(* IEC 61131-3 sources: 2026_Projet_YGO_ExcavatriceDragage/TOOLS/TEST_AUTO_CI/RESULTS/L_SIMULATION/reports, 11 files *)

(* ---- FB_Sim_Encoder_test.st ---- *)
(* =======================================================================
   Automated Unit Test - FB_Sim_Encoder
   ======================================================================= *)
TEST 'TC-P13-ENC-001 Enable FALSE conserve la valeur passee par VAR_IN_OUT'
VAR
    fb     : FB_Sim_Encoder;
    rawPos : UDINT := 1000;
END_VAR
    fb.Enable := FALSE;
    fb.StepNumber := 3;
    fb(RawPos := rawPos);
    ASSERT_EQ(fb.RawPosOut, 1000, 'Enable FALSE -> RawPosOut conserve la valeur persistee');
END_TEST

TEST 'TC-P13-ENC-002 Simulation incrementation comptage en montee'
VAR
    fb     : FB_Sim_Encoder;
    rawPos : UDINT := 1000;
    i      : INT;
END_VAR
    fb.Enable := TRUE;
    fb.RelayFwd := TRUE; (* Sens montee *)
    fb.RelayRev := FALSE;
    fb.StepNumber := 3;

    FOR i := 1 TO 10 DO
        fb(RawPos := rawPos);
    END_FOR;

    ASSERT_TRUE(fb.RawPosOut > 1000, 'RelayFwd TRUE -> RawPosOut augmente');
END_TEST

TEST 'TC-P13-034 SpeedReportTauS=0.0 conserve le saut instantane historique (non-regression)'
VAR
    fb     : FB_Sim_Encoder;
    rawPos : UDINT := 1000;
    i      : INT;
END_VAR
    fb.Enable := TRUE;
    fb.RelayFwd := TRUE;
    fb.StepNumber := 5;
    fb.SpeedReportTauS := 0.0;
    FOR i := 1 TO 5 DO
        fb(RawPos := rawPos);
    END_FOR;
    fb.RelayFwd := FALSE;
    fb.CoastDistanceM := 0.0;
    fb(RawPos := rawPos);
    ASSERT_EQ(fb.RawSpdOut, 0, 'Tau=0.0, coupure sans roulis -> vitesse rapportee tombe a 0 des le meme scan');
END_TEST

TEST 'TC-P13-035 SpeedReportTauS>0 fait decroitre RawSpdOut sur plusieurs scans (fidelite AX10, T316)'
VAR
    fb        : FB_Sim_Encoder;
    rawPos    : UDINT := 1000;
    i         : INT;
    spdAtCut  : DINT;
    spdNext   : DINT;
END_VAR
    fb.Enable := TRUE;
    fb.RelayFwd := TRUE;
    fb.StepNumber := 5;
    fb.SpeedReportTauS := 0.15; (* mirror tau M3 identifie sur trace, SYNTHETIQUE treuil *)
    fb.CoastDistanceM := 0.0;
    FOR i := 1 TO 20 DO
        fb(RawPos := rawPos); (* stabilise ReportedSpeedMps a la vitesse palier 5 *)
    END_FOR;
    fb.RelayFwd := FALSE;
    fb(RawPos := rawPos);
    spdAtCut := fb.RawSpdOut;
    fb(RawPos := rawPos);
    spdNext := fb.RawSpdOut;
    ASSERT_TRUE(spdAtCut > 0, 'Coupure relais : vitesse rapportee encore non nulle au 1er scan (pas de saut instantane)');
    ASSERT_TRUE(spdNext < spdAtCut, 'Vitesse rapportee decroit scan apres scan (rampe continue, pas un escalier)');
    ASSERT_TRUE(spdNext > 0, 'Decroissance progressive : pas encore a zero au 2e scan');
END_TEST

TEST 'TC-P13-031 PresetCmd applique PresetValue apres PresetLatencyCycles, mouvement gele pendant la latence'
VAR
    fb     : FB_Sim_Encoder;
    rawPos : UDINT := 1000;
END_VAR
    fb.Enable := TRUE;
    fb.RelayFwd := TRUE; (* commande de mouvement maintenue pendant le preset *)
    fb.StepNumber := 3;
    fb.PresetLatencyCycles := 2;
    fb.PresetValue := 500000;
    fb.PresetCmd := TRUE;
    fb(RawPos := rawPos);
    ASSERT_EQ(fb.RawPosOut, 1000, 'Pendant la latence : position brute conservee, mouvement gele');
    fb(RawPos := rawPos);
    ASSERT_EQ(fb.RawPosOut, 1000, 'Latence non ecoulee : position encore conservee');
    fb(RawPos := rawPos);
    ASSERT_EQ(fb.RawPosOut, 500000, 'Latence ecoulee : PresetValue charge (priorite sur Fwd/Rev)');
END_TEST

TEST 'TC-P13-032 Le comptage descend de facon continue et franchit 0 sans se figer (butee silencieuse supprimee)'
VAR
    fb        : FB_Sim_Encoder;
    rawPos    : UDINT := 41; (* 41 pts : exactement un pas de descente au palier 1 -> atteint 0 au 1er scan *)
    wrapAt41  : UDINT := 4294967255; (* 2^32 - 41 : -41 pts en representation signee 32 bits *)
    wrapAt82  : UDINT := 4294967214; (* 2^32 - 82 : -82 pts *)
END_VAR
    fb.Enable := TRUE;
    fb.RelayRev := TRUE;
    fb.StepNumber := 1; (* 1,0 m/s -> 1,0 x 4096 x 0,010 = 40,96 pts/scan, arrondi a 41 *)
    fb(RawPos := rawPos);
    rawPos := fb.RawPosOut; (* le caller conserve la memoire persistante du codeur *)
    ASSERT_EQ(fb.RawPosOut, 0, 'Un pas de descente amene le comptage exactement a 0 (point de passage)');
    fb(RawPos := rawPos);
    rawPos := fb.RawPosOut;
    ASSERT_TRUE(fb.RawPosOut <> 0, 'Scan suivant : le comptage franchit 0 au lieu de s y figer');
    ASSERT_EQ(fb.RawPosOut, wrapAt41, 'Comptage = -41 pts (aucune borne a 0)');
    fb(RawPos := rawPos);
    ASSERT_EQ(fb.RawPosOut, wrapAt82, 'Le comptage continue de decroitre : -82 pts');
END_TEST

TEST 'TC-P13-036 Comptage a 0 sous commande de descente : le scan suivant ne maintient pas 0'
VAR
    fb       : FB_Sim_Encoder;
    rawPos   : UDINT := 0; (* etat exact du blocage M2 du 2026-09-20 *)
    wrapAt41 : UDINT := 4294967255; (* 2^32 - 41 : -41 pts *)
END_VAR
    fb.Enable := TRUE;
    fb.RelayRev := TRUE;
    fb.StepNumber := 1;
    fb(RawPos := rawPos);
    rawPos := fb.RawPosOut;
    ASSERT_EQ(fb.RawPosOut, wrapAt41, 'Comptage a 0 + descente : passe a -41 pts, ne reste pas bloque a 0');
    fb(RawPos := rawPos);
    ASSERT_EQ(fb.RawPosOut, 4294967214, 'Le comptage poursuit sa descente au scan suivant (-82 pts)');
END_TEST

TEST 'TC-P13-037 Garde de plage : saturation signalee, comptage borne, aucune vitesse publiee'
VAR
    fb         : FB_Sim_Encoder;
    posLimit   : UDINT := 1073741824; (* +2^30 pts : limite de plage du modele *)
    negLimit   : UDINT := 3221225472; (* 2^32 - 2^30 : -2^30 pts en signe *)
END_VAR
    fb.Enable := TRUE;
    fb.RelayFwd := TRUE;
    fb.StepNumber := 5; (* palier 5 : 82 pts/scan *)
    fb(RawPos := posLimit);
    ASSERT_TRUE(fb.CountSaturated, 'Comptage hors plage haute : CountSaturated TRUE (saturation signalee)');
    ASSERT_EQ(fb.RawPosOut, posLimit, 'Comptage borne a la limite de plage (aucun rebouclage UDINT)');
    ASSERT_EQ(fb.RawSpdOut, 0, 'Position bornee : aucune vitesse de mouvement publiee (coherence)');
    fb.RelayFwd := FALSE;
    fb.RelayRev := TRUE;
    fb(RawPos := negLimit);
    ASSERT_TRUE(fb.CountSaturated, 'Comptage hors plage basse : CountSaturated TRUE');
    ASSERT_EQ(fb.RawPosOut, negLimit, 'Comptage borne a la limite basse (aucun rebouclage UDINT)');
    ASSERT_EQ(fb.RawSpdOut, 0, 'Saturation basse : vitesse de mouvement purge');
END_TEST

TEST 'TC-P13-038 Comptage negatif : la montee ramene vers 0 puis au-dela (continuite bidirectionnelle)'
VAR
    fb      : FB_Sim_Encoder;
    rawPos  : UDINT := 4294967255; (* 2^32 - 41 : -41 pts *)
END_VAR
    fb.Enable := TRUE;
    fb.RelayFwd := TRUE;
    fb.RelayRev := FALSE;
    fb.StepNumber := 1;
    fb(RawPos := rawPos);
    rawPos := fb.RawPosOut;
    ASSERT_EQ(fb.RawPosOut, 0, 'Depuis -41 pts : un pas de montee ramene exactement a 0');
    fb(RawPos := rawPos);
    ASSERT_EQ(fb.RawPosOut, 41, 'Le scan suivant poursuit au-dela de 0 (aucune butee dans les deux sens)');
END_TEST

(* ---- FB_Sim_Joystick_test.st ---- *)
(* =======================================================================
   Automated Unit Test - FB_Sim_Joystick
   ======================================================================= *)
TEST 'TC-P13-JOY-001 Enable FALSE -> positionne les axes au neutre (5000)'
VAR
    fb : FB_Sim_Joystick;
END_VAR
    fb.Enable := FALSE;
    fb();
    ASSERT_EQ(fb.RawX, 5000, 'Enable FALSE -> RawX au neutre NeutralRaw=5000');
    ASSERT_EQ(fb.RawY, 5000, 'Enable FALSE -> RawY au neutre NeutralRaw=5000');
    ASSERT_FALSE(fb.RawButton, 'Enable FALSE -> RawButton FALSE');
END_TEST

TEST 'TC-T418-001 Appui avant debattement puis relachement armement'
VAR
    fb : FB_Sim_Joystick;
    i  : INT;
END_VAR
    fb.Enable := TRUE;
    fb(); (* Relachement observe avant nouveau geste *)
    fb.BtnFwd_Up_Close := TRUE;
    fb();
    ASSERT_TRUE(fb.RawButton, 'Appui armement en premier');
    ASSERT_EQ(fb.RawY, 5000, 'Manche au neutre pendant appui');
    ADVANCE_TIME(10000000);
        fb();
ADVANCE_TIME(10000000);
        fb();
ADVANCE_TIME(10000000);
        fb();
ADVANCE_TIME(10000000);
        fb();
ADVANCE_TIME(10000000);
        fb();
ADVANCE_TIME(10000000);
        fb();
ADVANCE_TIME(10000000);
        fb();
ADVANCE_TIME(10000000);
        fb();
ADVANCE_TIME(10000000);
        fb();
ADVANCE_TIME(10000000);
        fb();
    ASSERT_TRUE(fb.RawButton, 'Appui tenu 100 ms');
    ASSERT_EQ(fb.RawY, 5000, 'Aucun debattement avant 200 ms');
    ADVANCE_TIME(10000000);
        fb();
ADVANCE_TIME(10000000);
        fb();
ADVANCE_TIME(10000000);
        fb();
ADVANCE_TIME(10000000);
        fb();
ADVANCE_TIME(10000000);
        fb();
ADVANCE_TIME(10000000);
        fb();
ADVANCE_TIME(10000000);
        fb();
ADVANCE_TIME(10000000);
        fb();
ADVANCE_TIME(10000000);
        fb();
ADVANCE_TIME(10000000);
        fb();
ADVANCE_TIME(10000000);
        fb();
ADVANCE_TIME(10000000);
        fb();
ADVANCE_TIME(10000000);
        fb();
ADVANCE_TIME(10000000);
        fb();
ADVANCE_TIME(10000000);
        fb();
ADVANCE_TIME(10000000);
        fb();
ADVANCE_TIME(10000000);
        fb();
ADVANCE_TIME(10000000);
        fb();
ADVANCE_TIME(10000000);
        fb();
ADVANCE_TIME(10000000);
        fb();
ADVANCE_TIME(10000000);
        fb();
ADVANCE_TIME(10000000);
        fb();
ADVANCE_TIME(10000000);
        fb();
ADVANCE_TIME(10000000);
        fb();
ADVANCE_TIME(10000000);
        fb();
    ASSERT_TRUE(fb.RawY > 5000, 'BtnFwd -> RawY monte vers MaxRaw');
    ASSERT_TRUE(fb.RawButton, 'Armement encore tenu au debut debattement');
    ADVANCE_TIME(10000000);
        fb();
        ASSERT_FALSE(fb.RawButton AND 1 > 20, 'Pas de nouvel appui apres relachement');
ADVANCE_TIME(10000000);
        fb();
        ASSERT_FALSE(fb.RawButton AND 2 > 20, 'Pas de nouvel appui apres relachement');
ADVANCE_TIME(10000000);
        fb();
        ASSERT_FALSE(fb.RawButton AND 3 > 20, 'Pas de nouvel appui apres relachement');
ADVANCE_TIME(10000000);
        fb();
        ASSERT_FALSE(fb.RawButton AND 4 > 20, 'Pas de nouvel appui apres relachement');
ADVANCE_TIME(10000000);
        fb();
        ASSERT_FALSE(fb.RawButton AND 5 > 20, 'Pas de nouvel appui apres relachement');
ADVANCE_TIME(10000000);
        fb();
        ASSERT_FALSE(fb.RawButton AND 6 > 20, 'Pas de nouvel appui apres relachement');
ADVANCE_TIME(10000000);
        fb();
        ASSERT_FALSE(fb.RawButton AND 7 > 20, 'Pas de nouvel appui apres relachement');
ADVANCE_TIME(10000000);
        fb();
        ASSERT_FALSE(fb.RawButton AND 8 > 20, 'Pas de nouvel appui apres relachement');
ADVANCE_TIME(10000000);
        fb();
        ASSERT_FALSE(fb.RawButton AND 9 > 20, 'Pas de nouvel appui apres relachement');
ADVANCE_TIME(10000000);
        fb();
        ASSERT_FALSE(fb.RawButton AND 10 > 20, 'Pas de nouvel appui apres relachement');
ADVANCE_TIME(10000000);
        fb();
        ASSERT_FALSE(fb.RawButton AND 11 > 20, 'Pas de nouvel appui apres relachement');
ADVANCE_TIME(10000000);
        fb();
        ASSERT_FALSE(fb.RawButton AND 12 > 20, 'Pas de nouvel appui apres relachement');
ADVANCE_TIME(10000000);
        fb();
        ASSERT_FALSE(fb.RawButton AND 13 > 20, 'Pas de nouvel appui apres relachement');
ADVANCE_TIME(10000000);
        fb();
        ASSERT_FALSE(fb.RawButton AND 14 > 20, 'Pas de nouvel appui apres relachement');
ADVANCE_TIME(10000000);
        fb();
        ASSERT_FALSE(fb.RawButton AND 15 > 20, 'Pas de nouvel appui apres relachement');
ADVANCE_TIME(10000000);
        fb();
        ASSERT_FALSE(fb.RawButton AND 16 > 20, 'Pas de nouvel appui apres relachement');
ADVANCE_TIME(10000000);
        fb();
        ASSERT_FALSE(fb.RawButton AND 17 > 20, 'Pas de nouvel appui apres relachement');
ADVANCE_TIME(10000000);
        fb();
        ASSERT_FALSE(fb.RawButton AND 18 > 20, 'Pas de nouvel appui apres relachement');
ADVANCE_TIME(10000000);
        fb();
        ASSERT_FALSE(fb.RawButton AND 19 > 20, 'Pas de nouvel appui apres relachement');
ADVANCE_TIME(10000000);
        fb();
        ASSERT_FALSE(fb.RawButton AND 20 > 20, 'Pas de nouvel appui apres relachement');
ADVANCE_TIME(10000000);
        fb();
        ASSERT_FALSE(fb.RawButton AND 21 > 20, 'Pas de nouvel appui apres relachement');
ADVANCE_TIME(10000000);
        fb();
        ASSERT_FALSE(fb.RawButton AND 22 > 20, 'Pas de nouvel appui apres relachement');
ADVANCE_TIME(10000000);
        fb();
        ASSERT_FALSE(fb.RawButton AND 23 > 20, 'Pas de nouvel appui apres relachement');
ADVANCE_TIME(10000000);
        fb();
        ASSERT_FALSE(fb.RawButton AND 24 > 20, 'Pas de nouvel appui apres relachement');
ADVANCE_TIME(10000000);
        fb();
        ASSERT_FALSE(fb.RawButton AND 25 > 20, 'Pas de nouvel appui apres relachement');
ADVANCE_TIME(10000000);
        fb();
        ASSERT_FALSE(fb.RawButton AND 26 > 20, 'Pas de nouvel appui apres relachement');
ADVANCE_TIME(10000000);
        fb();
        ASSERT_FALSE(fb.RawButton AND 27 > 20, 'Pas de nouvel appui apres relachement');
ADVANCE_TIME(10000000);
        fb();
        ASSERT_FALSE(fb.RawButton AND 28 > 20, 'Pas de nouvel appui apres relachement');
ADVANCE_TIME(10000000);
        fb();
        ASSERT_FALSE(fb.RawButton AND 29 > 20, 'Pas de nouvel appui apres relachement');
ADVANCE_TIME(10000000);
        fb();
        ASSERT_FALSE(fb.RawButton AND 30 > 20, 'Pas de nouvel appui apres relachement');
ADVANCE_TIME(10000000);
        fb();
        ASSERT_FALSE(fb.RawButton AND 31 > 20, 'Pas de nouvel appui apres relachement');
ADVANCE_TIME(10000000);
        fb();
        ASSERT_FALSE(fb.RawButton AND 32 > 20, 'Pas de nouvel appui apres relachement');
ADVANCE_TIME(10000000);
        fb();
        ASSERT_FALSE(fb.RawButton AND 33 > 20, 'Pas de nouvel appui apres relachement');
ADVANCE_TIME(10000000);
        fb();
        ASSERT_FALSE(fb.RawButton AND 34 > 20, 'Pas de nouvel appui apres relachement');
ADVANCE_TIME(10000000);
        fb();
        ASSERT_FALSE(fb.RawButton AND 35 > 20, 'Pas de nouvel appui apres relachement');
ADVANCE_TIME(10000000);
        fb();
        ASSERT_FALSE(fb.RawButton AND 36 > 20, 'Pas de nouvel appui apres relachement');
ADVANCE_TIME(10000000);
        fb();
        ASSERT_FALSE(fb.RawButton AND 37 > 20, 'Pas de nouvel appui apres relachement');
ADVANCE_TIME(10000000);
        fb();
        ASSERT_FALSE(fb.RawButton AND 38 > 20, 'Pas de nouvel appui apres relachement');
ADVANCE_TIME(10000000);
        fb();
        ASSERT_FALSE(fb.RawButton AND 39 > 20, 'Pas de nouvel appui apres relachement');
ADVANCE_TIME(10000000);
        fb();
        ASSERT_FALSE(fb.RawButton AND 40 > 20, 'Pas de nouvel appui apres relachement');
ADVANCE_TIME(10000000);
        fb();
        ASSERT_FALSE(fb.RawButton AND 41 > 20, 'Pas de nouvel appui apres relachement');
ADVANCE_TIME(10000000);
        fb();
        ASSERT_FALSE(fb.RawButton AND 42 > 20, 'Pas de nouvel appui apres relachement');
ADVANCE_TIME(10000000);
        fb();
        ASSERT_FALSE(fb.RawButton AND 43 > 20, 'Pas de nouvel appui apres relachement');
ADVANCE_TIME(10000000);
        fb();
        ASSERT_FALSE(fb.RawButton AND 44 > 20, 'Pas de nouvel appui apres relachement');
ADVANCE_TIME(10000000);
        fb();
        ASSERT_FALSE(fb.RawButton AND 45 > 20, 'Pas de nouvel appui apres relachement');
ADVANCE_TIME(10000000);
        fb();
        ASSERT_FALSE(fb.RawButton AND 46 > 20, 'Pas de nouvel appui apres relachement');
ADVANCE_TIME(10000000);
        fb();
        ASSERT_FALSE(fb.RawButton AND 47 > 20, 'Pas de nouvel appui apres relachement');
ADVANCE_TIME(10000000);
        fb();
        ASSERT_FALSE(fb.RawButton AND 48 > 20, 'Pas de nouvel appui apres relachement');
ADVANCE_TIME(10000000);
        fb();
        ASSERT_FALSE(fb.RawButton AND 49 > 20, 'Pas de nouvel appui apres relachement');
ADVANCE_TIME(10000000);
        fb();
        ASSERT_FALSE(fb.RawButton AND 50 > 20, 'Pas de nouvel appui apres relachement');
ADVANCE_TIME(10000000);
        fb();
        ASSERT_FALSE(fb.RawButton AND 51 > 20, 'Pas de nouvel appui apres relachement');
ADVANCE_TIME(10000000);
        fb();
        ASSERT_FALSE(fb.RawButton AND 52 > 20, 'Pas de nouvel appui apres relachement');
ADVANCE_TIME(10000000);
        fb();
        ASSERT_FALSE(fb.RawButton AND 53 > 20, 'Pas de nouvel appui apres relachement');
ADVANCE_TIME(10000000);
        fb();
        ASSERT_FALSE(fb.RawButton AND 54 > 20, 'Pas de nouvel appui apres relachement');
ADVANCE_TIME(10000000);
        fb();
        ASSERT_FALSE(fb.RawButton AND 55 > 20, 'Pas de nouvel appui apres relachement');
ADVANCE_TIME(10000000);
        fb();
        ASSERT_FALSE(fb.RawButton AND 56 > 20, 'Pas de nouvel appui apres relachement');
ADVANCE_TIME(10000000);
        fb();
        ASSERT_FALSE(fb.RawButton AND 57 > 20, 'Pas de nouvel appui apres relachement');
ADVANCE_TIME(10000000);
        fb();
        ASSERT_FALSE(fb.RawButton AND 58 > 20, 'Pas de nouvel appui apres relachement');
ADVANCE_TIME(10000000);
        fb();
        ASSERT_FALSE(fb.RawButton AND 59 > 20, 'Pas de nouvel appui apres relachement');
ADVANCE_TIME(10000000);
        fb();
        ASSERT_FALSE(fb.RawButton AND 60 > 20, 'Pas de nouvel appui apres relachement');
ADVANCE_TIME(10000000);
        fb();
        ASSERT_FALSE(fb.RawButton AND 61 > 20, 'Pas de nouvel appui apres relachement');
ADVANCE_TIME(10000000);
        fb();
        ASSERT_FALSE(fb.RawButton AND 62 > 20, 'Pas de nouvel appui apres relachement');
ADVANCE_TIME(10000000);
        fb();
        ASSERT_FALSE(fb.RawButton AND 63 > 20, 'Pas de nouvel appui apres relachement');
ADVANCE_TIME(10000000);
        fb();
        ASSERT_FALSE(fb.RawButton AND 64 > 20, 'Pas de nouvel appui apres relachement');
ADVANCE_TIME(10000000);
        fb();
        ASSERT_FALSE(fb.RawButton AND 65 > 20, 'Pas de nouvel appui apres relachement');
ADVANCE_TIME(10000000);
        fb();
        ASSERT_FALSE(fb.RawButton AND 66 > 20, 'Pas de nouvel appui apres relachement');
ADVANCE_TIME(10000000);
        fb();
        ASSERT_FALSE(fb.RawButton AND 67 > 20, 'Pas de nouvel appui apres relachement');
ADVANCE_TIME(10000000);
        fb();
        ASSERT_FALSE(fb.RawButton AND 68 > 20, 'Pas de nouvel appui apres relachement');
ADVANCE_TIME(10000000);
        fb();
        ASSERT_FALSE(fb.RawButton AND 69 > 20, 'Pas de nouvel appui apres relachement');
ADVANCE_TIME(10000000);
        fb();
        ASSERT_FALSE(fb.RawButton AND 70 > 20, 'Pas de nouvel appui apres relachement');
ADVANCE_TIME(10000000);
        fb();
        ASSERT_FALSE(fb.RawButton AND 71 > 20, 'Pas de nouvel appui apres relachement');
ADVANCE_TIME(10000000);
        fb();
        ASSERT_FALSE(fb.RawButton AND 72 > 20, 'Pas de nouvel appui apres relachement');
ADVANCE_TIME(10000000);
        fb();
        ASSERT_FALSE(fb.RawButton AND 73 > 20, 'Pas de nouvel appui apres relachement');
ADVANCE_TIME(10000000);
        fb();
        ASSERT_FALSE(fb.RawButton AND 74 > 20, 'Pas de nouvel appui apres relachement');
ADVANCE_TIME(10000000);
        fb();
        ASSERT_FALSE(fb.RawButton AND 75 > 20, 'Pas de nouvel appui apres relachement');
ADVANCE_TIME(10000000);
        fb();
        ASSERT_FALSE(fb.RawButton AND 76 > 20, 'Pas de nouvel appui apres relachement');
ADVANCE_TIME(10000000);
        fb();
        ASSERT_FALSE(fb.RawButton AND 77 > 20, 'Pas de nouvel appui apres relachement');
ADVANCE_TIME(10000000);
        fb();
        ASSERT_FALSE(fb.RawButton AND 78 > 20, 'Pas de nouvel appui apres relachement');
ADVANCE_TIME(10000000);
        fb();
        ASSERT_FALSE(fb.RawButton AND 79 > 20, 'Pas de nouvel appui apres relachement');
ADVANCE_TIME(10000000);
        fb();
        ASSERT_FALSE(fb.RawButton AND 80 > 20, 'Pas de nouvel appui apres relachement');
ADVANCE_TIME(10000000);
        fb();
        ASSERT_FALSE(fb.RawButton AND 81 > 20, 'Pas de nouvel appui apres relachement');
ADVANCE_TIME(10000000);
        fb();
        ASSERT_FALSE(fb.RawButton AND 82 > 20, 'Pas de nouvel appui apres relachement');
ADVANCE_TIME(10000000);
        fb();
        ASSERT_FALSE(fb.RawButton AND 83 > 20, 'Pas de nouvel appui apres relachement');
ADVANCE_TIME(10000000);
        fb();
        ASSERT_FALSE(fb.RawButton AND 84 > 20, 'Pas de nouvel appui apres relachement');
ADVANCE_TIME(10000000);
        fb();
        ASSERT_FALSE(fb.RawButton AND 85 > 20, 'Pas de nouvel appui apres relachement');
ADVANCE_TIME(10000000);
        fb();
        ASSERT_FALSE(fb.RawButton AND 86 > 20, 'Pas de nouvel appui apres relachement');
ADVANCE_TIME(10000000);
        fb();
        ASSERT_FALSE(fb.RawButton AND 87 > 20, 'Pas de nouvel appui apres relachement');
ADVANCE_TIME(10000000);
        fb();
        ASSERT_FALSE(fb.RawButton AND 88 > 20, 'Pas de nouvel appui apres relachement');
ADVANCE_TIME(10000000);
        fb();
        ASSERT_FALSE(fb.RawButton AND 89 > 20, 'Pas de nouvel appui apres relachement');
ADVANCE_TIME(10000000);
        fb();
        ASSERT_FALSE(fb.RawButton AND 90 > 20, 'Pas de nouvel appui apres relachement');
ADVANCE_TIME(10000000);
        fb();
        ASSERT_FALSE(fb.RawButton AND 91 > 20, 'Pas de nouvel appui apres relachement');
ADVANCE_TIME(10000000);
        fb();
        ASSERT_FALSE(fb.RawButton AND 92 > 20, 'Pas de nouvel appui apres relachement');
ADVANCE_TIME(10000000);
        fb();
        ASSERT_FALSE(fb.RawButton AND 93 > 20, 'Pas de nouvel appui apres relachement');
ADVANCE_TIME(10000000);
        fb();
        ASSERT_FALSE(fb.RawButton AND 94 > 20, 'Pas de nouvel appui apres relachement');
ADVANCE_TIME(10000000);
        fb();
        ASSERT_FALSE(fb.RawButton AND 95 > 20, 'Pas de nouvel appui apres relachement');
ADVANCE_TIME(10000000);
        fb();
        ASSERT_FALSE(fb.RawButton AND 96 > 20, 'Pas de nouvel appui apres relachement');
ADVANCE_TIME(10000000);
        fb();
        ASSERT_FALSE(fb.RawButton AND 97 > 20, 'Pas de nouvel appui apres relachement');
ADVANCE_TIME(10000000);
        fb();
        ASSERT_FALSE(fb.RawButton AND 98 > 20, 'Pas de nouvel appui apres relachement');
ADVANCE_TIME(10000000);
        fb();
        ASSERT_FALSE(fb.RawButton AND 99 > 20, 'Pas de nouvel appui apres relachement');
ADVANCE_TIME(10000000);
        fb();
        ASSERT_FALSE(fb.RawButton AND 100 > 20, 'Pas de nouvel appui apres relachement');
ADVANCE_TIME(10000000);
        fb();
        ASSERT_FALSE(fb.RawButton AND 101 > 20, 'Pas de nouvel appui apres relachement');
ADVANCE_TIME(10000000);
        fb();
        ASSERT_FALSE(fb.RawButton AND 102 > 20, 'Pas de nouvel appui apres relachement');
ADVANCE_TIME(10000000);
        fb();
        ASSERT_FALSE(fb.RawButton AND 103 > 20, 'Pas de nouvel appui apres relachement');
ADVANCE_TIME(10000000);
        fb();
        ASSERT_FALSE(fb.RawButton AND 104 > 20, 'Pas de nouvel appui apres relachement');
ADVANCE_TIME(10000000);
        fb();
        ASSERT_FALSE(fb.RawButton AND 105 > 20, 'Pas de nouvel appui apres relachement');
ADVANCE_TIME(10000000);
        fb();
        ASSERT_FALSE(fb.RawButton AND 106 > 20, 'Pas de nouvel appui apres relachement');
ADVANCE_TIME(10000000);
        fb();
        ASSERT_FALSE(fb.RawButton AND 107 > 20, 'Pas de nouvel appui apres relachement');
ADVANCE_TIME(10000000);
        fb();
        ASSERT_FALSE(fb.RawButton AND 108 > 20, 'Pas de nouvel appui apres relachement');
ADVANCE_TIME(10000000);
        fb();
        ASSERT_FALSE(fb.RawButton AND 109 > 20, 'Pas de nouvel appui apres relachement');
ADVANCE_TIME(10000000);
        fb();
        ASSERT_FALSE(fb.RawButton AND 110 > 20, 'Pas de nouvel appui apres relachement');
ADVANCE_TIME(10000000);
        fb();
        ASSERT_FALSE(fb.RawButton AND 111 > 20, 'Pas de nouvel appui apres relachement');
ADVANCE_TIME(10000000);
        fb();
        ASSERT_FALSE(fb.RawButton AND 112 > 20, 'Pas de nouvel appui apres relachement');
ADVANCE_TIME(10000000);
        fb();
        ASSERT_FALSE(fb.RawButton AND 113 > 20, 'Pas de nouvel appui apres relachement');
ADVANCE_TIME(10000000);
        fb();
        ASSERT_FALSE(fb.RawButton AND 114 > 20, 'Pas de nouvel appui apres relachement');
ADVANCE_TIME(10000000);
        fb();
        ASSERT_FALSE(fb.RawButton AND 115 > 20, 'Pas de nouvel appui apres relachement');
ADVANCE_TIME(10000000);
        fb();
        ASSERT_FALSE(fb.RawButton AND 116 > 20, 'Pas de nouvel appui apres relachement');
ADVANCE_TIME(10000000);
        fb();
        ASSERT_FALSE(fb.RawButton AND 117 > 20, 'Pas de nouvel appui apres relachement');
ADVANCE_TIME(10000000);
        fb();
        ASSERT_FALSE(fb.RawButton AND 118 > 20, 'Pas de nouvel appui apres relachement');
ADVANCE_TIME(10000000);
        fb();
        ASSERT_FALSE(fb.RawButton AND 119 > 20, 'Pas de nouvel appui apres relachement');
ADVANCE_TIME(10000000);
        fb();
        ASSERT_FALSE(fb.RawButton AND 120 > 20, 'Pas de nouvel appui apres relachement');
ADVANCE_TIME(10000000);
        fb();
        ASSERT_FALSE(fb.RawButton AND 121 > 20, 'Pas de nouvel appui apres relachement');
ADVANCE_TIME(10000000);
        fb();
        ASSERT_FALSE(fb.RawButton AND 122 > 20, 'Pas de nouvel appui apres relachement');
ADVANCE_TIME(10000000);
        fb();
        ASSERT_FALSE(fb.RawButton AND 123 > 20, 'Pas de nouvel appui apres relachement');
ADVANCE_TIME(10000000);
        fb();
        ASSERT_FALSE(fb.RawButton AND 124 > 20, 'Pas de nouvel appui apres relachement');
ADVANCE_TIME(10000000);
        fb();
        ASSERT_FALSE(fb.RawButton AND 125 > 20, 'Pas de nouvel appui apres relachement');
ADVANCE_TIME(10000000);
        fb();
        ASSERT_FALSE(fb.RawButton AND 126 > 20, 'Pas de nouvel appui apres relachement');
ADVANCE_TIME(10000000);
        fb();
        ASSERT_FALSE(fb.RawButton AND 127 > 20, 'Pas de nouvel appui apres relachement');
ADVANCE_TIME(10000000);
        fb();
        ASSERT_FALSE(fb.RawButton AND 128 > 20, 'Pas de nouvel appui apres relachement');
ADVANCE_TIME(10000000);
        fb();
        ASSERT_FALSE(fb.RawButton AND 129 > 20, 'Pas de nouvel appui apres relachement');
ADVANCE_TIME(10000000);
        fb();
        ASSERT_FALSE(fb.RawButton AND 130 > 20, 'Pas de nouvel appui apres relachement');
ADVANCE_TIME(10000000);
        fb();
        ASSERT_FALSE(fb.RawButton AND 131 > 20, 'Pas de nouvel appui apres relachement');
ADVANCE_TIME(10000000);
        fb();
        ASSERT_FALSE(fb.RawButton AND 132 > 20, 'Pas de nouvel appui apres relachement');
ADVANCE_TIME(10000000);
        fb();
        ASSERT_FALSE(fb.RawButton AND 133 > 20, 'Pas de nouvel appui apres relachement');
ADVANCE_TIME(10000000);
        fb();
        ASSERT_FALSE(fb.RawButton AND 134 > 20, 'Pas de nouvel appui apres relachement');
ADVANCE_TIME(10000000);
        fb();
        ASSERT_FALSE(fb.RawButton AND 135 > 20, 'Pas de nouvel appui apres relachement');
ADVANCE_TIME(10000000);
        fb();
        ASSERT_FALSE(fb.RawButton AND 136 > 20, 'Pas de nouvel appui apres relachement');
ADVANCE_TIME(10000000);
        fb();
        ASSERT_FALSE(fb.RawButton AND 137 > 20, 'Pas de nouvel appui apres relachement');
ADVANCE_TIME(10000000);
        fb();
        ASSERT_FALSE(fb.RawButton AND 138 > 20, 'Pas de nouvel appui apres relachement');
ADVANCE_TIME(10000000);
        fb();
        ASSERT_FALSE(fb.RawButton AND 139 > 20, 'Pas de nouvel appui apres relachement');
ADVANCE_TIME(10000000);
        fb();
        ASSERT_FALSE(fb.RawButton AND 140 > 20, 'Pas de nouvel appui apres relachement');
ADVANCE_TIME(10000000);
        fb();
        ASSERT_FALSE(fb.RawButton AND 141 > 20, 'Pas de nouvel appui apres relachement');
ADVANCE_TIME(10000000);
        fb();
        ASSERT_FALSE(fb.RawButton AND 142 > 20, 'Pas de nouvel appui apres relachement');
ADVANCE_TIME(10000000);
        fb();
        ASSERT_FALSE(fb.RawButton AND 143 > 20, 'Pas de nouvel appui apres relachement');
ADVANCE_TIME(10000000);
        fb();
        ASSERT_FALSE(fb.RawButton AND 144 > 20, 'Pas de nouvel appui apres relachement');
ADVANCE_TIME(10000000);
        fb();
        ASSERT_FALSE(fb.RawButton AND 145 > 20, 'Pas de nouvel appui apres relachement');
ADVANCE_TIME(10000000);
        fb();
        ASSERT_FALSE(fb.RawButton AND 146 > 20, 'Pas de nouvel appui apres relachement');
ADVANCE_TIME(10000000);
        fb();
        ASSERT_FALSE(fb.RawButton AND 147 > 20, 'Pas de nouvel appui apres relachement');
ADVANCE_TIME(10000000);
        fb();
        ASSERT_FALSE(fb.RawButton AND 148 > 20, 'Pas de nouvel appui apres relachement');
ADVANCE_TIME(10000000);
        fb();
        ASSERT_FALSE(fb.RawButton AND 149 > 20, 'Pas de nouvel appui apres relachement');
ADVANCE_TIME(10000000);
        fb();
        ASSERT_FALSE(fb.RawButton AND 150 > 20, 'Pas de nouvel appui apres relachement');
ADVANCE_TIME(10000000);
        fb();
        ASSERT_FALSE(fb.RawButton AND 151 > 20, 'Pas de nouvel appui apres relachement');
ADVANCE_TIME(10000000);
        fb();
        ASSERT_FALSE(fb.RawButton AND 152 > 20, 'Pas de nouvel appui apres relachement');
ADVANCE_TIME(10000000);
        fb();
        ASSERT_FALSE(fb.RawButton AND 153 > 20, 'Pas de nouvel appui apres relachement');
ADVANCE_TIME(10000000);
        fb();
        ASSERT_FALSE(fb.RawButton AND 154 > 20, 'Pas de nouvel appui apres relachement');
ADVANCE_TIME(10000000);
        fb();
        ASSERT_FALSE(fb.RawButton AND 155 > 20, 'Pas de nouvel appui apres relachement');
ADVANCE_TIME(10000000);
        fb();
        ASSERT_FALSE(fb.RawButton AND 156 > 20, 'Pas de nouvel appui apres relachement');
ADVANCE_TIME(10000000);
        fb();
        ASSERT_FALSE(fb.RawButton AND 157 > 20, 'Pas de nouvel appui apres relachement');
ADVANCE_TIME(10000000);
        fb();
        ASSERT_FALSE(fb.RawButton AND 158 > 20, 'Pas de nouvel appui apres relachement');
ADVANCE_TIME(10000000);
        fb();
        ASSERT_FALSE(fb.RawButton AND 159 > 20, 'Pas de nouvel appui apres relachement');
ADVANCE_TIME(10000000);
        fb();
        ASSERT_FALSE(fb.RawButton AND 160 > 20, 'Pas de nouvel appui apres relachement');
ADVANCE_TIME(10000000);
        fb();
        ASSERT_FALSE(fb.RawButton AND 161 > 20, 'Pas de nouvel appui apres relachement');
ADVANCE_TIME(10000000);
        fb();
        ASSERT_FALSE(fb.RawButton AND 162 > 20, 'Pas de nouvel appui apres relachement');
ADVANCE_TIME(10000000);
        fb();
        ASSERT_FALSE(fb.RawButton AND 163 > 20, 'Pas de nouvel appui apres relachement');
ADVANCE_TIME(10000000);
        fb();
        ASSERT_FALSE(fb.RawButton AND 164 > 20, 'Pas de nouvel appui apres relachement');
ADVANCE_TIME(10000000);
        fb();
        ASSERT_FALSE(fb.RawButton AND 165 > 20, 'Pas de nouvel appui apres relachement');
ADVANCE_TIME(10000000);
        fb();
        ASSERT_FALSE(fb.RawButton AND 166 > 20, 'Pas de nouvel appui apres relachement');
ADVANCE_TIME(10000000);
        fb();
        ASSERT_FALSE(fb.RawButton AND 167 > 20, 'Pas de nouvel appui apres relachement');
ADVANCE_TIME(10000000);
        fb();
        ASSERT_FALSE(fb.RawButton AND 168 > 20, 'Pas de nouvel appui apres relachement');
ADVANCE_TIME(10000000);
        fb();
        ASSERT_FALSE(fb.RawButton AND 169 > 20, 'Pas de nouvel appui apres relachement');
ADVANCE_TIME(10000000);
        fb();
        ASSERT_FALSE(fb.RawButton AND 170 > 20, 'Pas de nouvel appui apres relachement');
ADVANCE_TIME(10000000);
        fb();
        ASSERT_FALSE(fb.RawButton AND 171 > 20, 'Pas de nouvel appui apres relachement');
ADVANCE_TIME(10000000);
        fb();
        ASSERT_FALSE(fb.RawButton AND 172 > 20, 'Pas de nouvel appui apres relachement');
ADVANCE_TIME(10000000);
        fb();
        ASSERT_FALSE(fb.RawButton AND 173 > 20, 'Pas de nouvel appui apres relachement');
ADVANCE_TIME(10000000);
        fb();
        ASSERT_FALSE(fb.RawButton AND 174 > 20, 'Pas de nouvel appui apres relachement');
ADVANCE_TIME(10000000);
        fb();
        ASSERT_FALSE(fb.RawButton AND 175 > 20, 'Pas de nouvel appui apres relachement');
ADVANCE_TIME(10000000);
        fb();
        ASSERT_FALSE(fb.RawButton AND 176 > 20, 'Pas de nouvel appui apres relachement');
ADVANCE_TIME(10000000);
        fb();
        ASSERT_FALSE(fb.RawButton AND 177 > 20, 'Pas de nouvel appui apres relachement');
ADVANCE_TIME(10000000);
        fb();
        ASSERT_FALSE(fb.RawButton AND 178 > 20, 'Pas de nouvel appui apres relachement');
ADVANCE_TIME(10000000);
        fb();
        ASSERT_FALSE(fb.RawButton AND 179 > 20, 'Pas de nouvel appui apres relachement');
ADVANCE_TIME(10000000);
        fb();
        ASSERT_FALSE(fb.RawButton AND 180 > 20, 'Pas de nouvel appui apres relachement');
ADVANCE_TIME(10000000);
        fb();
        ASSERT_FALSE(fb.RawButton AND 181 > 20, 'Pas de nouvel appui apres relachement');
ADVANCE_TIME(10000000);
        fb();
        ASSERT_FALSE(fb.RawButton AND 182 > 20, 'Pas de nouvel appui apres relachement');
ADVANCE_TIME(10000000);
        fb();
        ASSERT_FALSE(fb.RawButton AND 183 > 20, 'Pas de nouvel appui apres relachement');
ADVANCE_TIME(10000000);
        fb();
        ASSERT_FALSE(fb.RawButton AND 184 > 20, 'Pas de nouvel appui apres relachement');
ADVANCE_TIME(10000000);
        fb();
        ASSERT_FALSE(fb.RawButton AND 185 > 20, 'Pas de nouvel appui apres relachement');
ADVANCE_TIME(10000000);
        fb();
        ASSERT_FALSE(fb.RawButton AND 186 > 20, 'Pas de nouvel appui apres relachement');
ADVANCE_TIME(10000000);
        fb();
        ASSERT_FALSE(fb.RawButton AND 187 > 20, 'Pas de nouvel appui apres relachement');
ADVANCE_TIME(10000000);
        fb();
        ASSERT_FALSE(fb.RawButton AND 188 > 20, 'Pas de nouvel appui apres relachement');
ADVANCE_TIME(10000000);
        fb();
        ASSERT_FALSE(fb.RawButton AND 189 > 20, 'Pas de nouvel appui apres relachement');
ADVANCE_TIME(10000000);
        fb();
        ASSERT_FALSE(fb.RawButton AND 190 > 20, 'Pas de nouvel appui apres relachement');
ADVANCE_TIME(10000000);
        fb();
        ASSERT_FALSE(fb.RawButton AND 191 > 20, 'Pas de nouvel appui apres relachement');
ADVANCE_TIME(10000000);
        fb();
        ASSERT_FALSE(fb.RawButton AND 192 > 20, 'Pas de nouvel appui apres relachement');
ADVANCE_TIME(10000000);
        fb();
        ASSERT_FALSE(fb.RawButton AND 193 > 20, 'Pas de nouvel appui apres relachement');
ADVANCE_TIME(10000000);
        fb();
        ASSERT_FALSE(fb.RawButton AND 194 > 20, 'Pas de nouvel appui apres relachement');
ADVANCE_TIME(10000000);
        fb();
        ASSERT_FALSE(fb.RawButton AND 195 > 20, 'Pas de nouvel appui apres relachement');
ADVANCE_TIME(10000000);
        fb();
        ASSERT_FALSE(fb.RawButton AND 196 > 20, 'Pas de nouvel appui apres relachement');
ADVANCE_TIME(10000000);
        fb();
        ASSERT_FALSE(fb.RawButton AND 197 > 20, 'Pas de nouvel appui apres relachement');
ADVANCE_TIME(10000000);
        fb();
        ASSERT_FALSE(fb.RawButton AND 198 > 20, 'Pas de nouvel appui apres relachement');
ADVANCE_TIME(10000000);
        fb();
        ASSERT_FALSE(fb.RawButton AND 199 > 20, 'Pas de nouvel appui apres relachement');
ADVANCE_TIME(10000000);
        fb();
        ASSERT_FALSE(fb.RawButton AND 200 > 20, 'Pas de nouvel appui apres relachement');
ADVANCE_TIME(10000000);
        fb();
        ASSERT_FALSE(fb.RawButton AND 201 > 20, 'Pas de nouvel appui apres relachement');
ADVANCE_TIME(10000000);
        fb();
        ASSERT_FALSE(fb.RawButton AND 202 > 20, 'Pas de nouvel appui apres relachement');
ADVANCE_TIME(10000000);
        fb();
        ASSERT_FALSE(fb.RawButton AND 203 > 20, 'Pas de nouvel appui apres relachement');
ADVANCE_TIME(10000000);
        fb();
        ASSERT_FALSE(fb.RawButton AND 204 > 20, 'Pas de nouvel appui apres relachement');
ADVANCE_TIME(10000000);
        fb();
        ASSERT_FALSE(fb.RawButton AND 205 > 20, 'Pas de nouvel appui apres relachement');
ADVANCE_TIME(10000000);
        fb();
        ASSERT_FALSE(fb.RawButton AND 206 > 20, 'Pas de nouvel appui apres relachement');
ADVANCE_TIME(10000000);
        fb();
        ASSERT_FALSE(fb.RawButton AND 207 > 20, 'Pas de nouvel appui apres relachement');
ADVANCE_TIME(10000000);
        fb();
        ASSERT_FALSE(fb.RawButton AND 208 > 20, 'Pas de nouvel appui apres relachement');
ADVANCE_TIME(10000000);
        fb();
        ASSERT_FALSE(fb.RawButton AND 209 > 20, 'Pas de nouvel appui apres relachement');
ADVANCE_TIME(10000000);
        fb();
        ASSERT_FALSE(fb.RawButton AND 210 > 20, 'Pas de nouvel appui apres relachement');
ADVANCE_TIME(10000000);
        fb();
        ASSERT_FALSE(fb.RawButton AND 211 > 20, 'Pas de nouvel appui apres relachement');
ADVANCE_TIME(10000000);
        fb();
        ASSERT_FALSE(fb.RawButton AND 212 > 20, 'Pas de nouvel appui apres relachement');
ADVANCE_TIME(10000000);
        fb();
        ASSERT_FALSE(fb.RawButton AND 213 > 20, 'Pas de nouvel appui apres relachement');
ADVANCE_TIME(10000000);
        fb();
        ASSERT_FALSE(fb.RawButton AND 214 > 20, 'Pas de nouvel appui apres relachement');
ADVANCE_TIME(10000000);
        fb();
        ASSERT_FALSE(fb.RawButton AND 215 > 20, 'Pas de nouvel appui apres relachement');
ADVANCE_TIME(10000000);
        fb();
        ASSERT_FALSE(fb.RawButton AND 216 > 20, 'Pas de nouvel appui apres relachement');
ADVANCE_TIME(10000000);
        fb();
        ASSERT_FALSE(fb.RawButton AND 217 > 20, 'Pas de nouvel appui apres relachement');
ADVANCE_TIME(10000000);
        fb();
        ASSERT_FALSE(fb.RawButton AND 218 > 20, 'Pas de nouvel appui apres relachement');
ADVANCE_TIME(10000000);
        fb();
        ASSERT_FALSE(fb.RawButton AND 219 > 20, 'Pas de nouvel appui apres relachement');
ADVANCE_TIME(10000000);
        fb();
        ASSERT_FALSE(fb.RawButton AND 220 > 20, 'Pas de nouvel appui apres relachement');
    ASSERT_FALSE(fb.RawButton, 'Bouton armement relache malgre maintien IHM');
    ASSERT_TRUE(fb.RawY > 9000, 'Manche reste deplace');
    fb.BtnFwd_Up_Close := FALSE;
    ADVANCE_TIME(10000000);
        fb();
ADVANCE_TIME(10000000);
        fb();
ADVANCE_TIME(10000000);
        fb();
ADVANCE_TIME(10000000);
        fb();
ADVANCE_TIME(10000000);
        fb();
ADVANCE_TIME(10000000);
        fb();
ADVANCE_TIME(10000000);
        fb();
ADVANCE_TIME(10000000);
        fb();
ADVANCE_TIME(10000000);
        fb();
ADVANCE_TIME(10000000);
        fb();
ADVANCE_TIME(10000000);
        fb();
ADVANCE_TIME(10000000);
        fb();
ADVANCE_TIME(10000000);
        fb();
ADVANCE_TIME(10000000);
        fb();
ADVANCE_TIME(10000000);
        fb();
ADVANCE_TIME(10000000);
        fb();
ADVANCE_TIME(10000000);
        fb();
ADVANCE_TIME(10000000);
        fb();
ADVANCE_TIME(10000000);
        fb();
ADVANCE_TIME(10000000);
        fb();
ADVANCE_TIME(10000000);
        fb();
ADVANCE_TIME(10000000);
        fb();
ADVANCE_TIME(10000000);
        fb();
ADVANCE_TIME(10000000);
        fb();
ADVANCE_TIME(10000000);
        fb();
ADVANCE_TIME(10000000);
        fb();
ADVANCE_TIME(10000000);
        fb();
ADVANCE_TIME(10000000);
        fb();
ADVANCE_TIME(10000000);
        fb();
ADVANCE_TIME(10000000);
        fb();
    ASSERT_EQ(fb.RawY, 5000, 'Retour au neutre au relachement IHM');
    ASSERT_FALSE(fb.ModelActive, 'Fin de propriete automatique');
END_TEST

TEST 'TC-T418-002 Bouton deja tenu au demarrage ou reactivation'
VAR
    fb : FB_Sim_Joystick;
    i : INT;
END_VAR
    fb.Enable := TRUE; fb.BtnRight_Fwd_MAINT := TRUE;
    ADVANCE_TIME(10000000); fb();
        ASSERT_FALSE(fb.RawButton, 'Demarrage tenu ne simule aucun appui');
        ASSERT_EQ(fb.RawX, 5000, 'Demarrage tenu neutre');
ADVANCE_TIME(10000000); fb();
        ASSERT_FALSE(fb.RawButton, 'Demarrage tenu ne simule aucun appui');
        ASSERT_EQ(fb.RawX, 5000, 'Demarrage tenu neutre');
ADVANCE_TIME(10000000); fb();
        ASSERT_FALSE(fb.RawButton, 'Demarrage tenu ne simule aucun appui');
        ASSERT_EQ(fb.RawX, 5000, 'Demarrage tenu neutre');
ADVANCE_TIME(10000000); fb();
        ASSERT_FALSE(fb.RawButton, 'Demarrage tenu ne simule aucun appui');
        ASSERT_EQ(fb.RawX, 5000, 'Demarrage tenu neutre');
ADVANCE_TIME(10000000); fb();
        ASSERT_FALSE(fb.RawButton, 'Demarrage tenu ne simule aucun appui');
        ASSERT_EQ(fb.RawX, 5000, 'Demarrage tenu neutre');
ADVANCE_TIME(10000000); fb();
        ASSERT_FALSE(fb.RawButton, 'Demarrage tenu ne simule aucun appui');
        ASSERT_EQ(fb.RawX, 5000, 'Demarrage tenu neutre');
ADVANCE_TIME(10000000); fb();
        ASSERT_FALSE(fb.RawButton, 'Demarrage tenu ne simule aucun appui');
        ASSERT_EQ(fb.RawX, 5000, 'Demarrage tenu neutre');
ADVANCE_TIME(10000000); fb();
        ASSERT_FALSE(fb.RawButton, 'Demarrage tenu ne simule aucun appui');
        ASSERT_EQ(fb.RawX, 5000, 'Demarrage tenu neutre');
ADVANCE_TIME(10000000); fb();
        ASSERT_FALSE(fb.RawButton, 'Demarrage tenu ne simule aucun appui');
        ASSERT_EQ(fb.RawX, 5000, 'Demarrage tenu neutre');
ADVANCE_TIME(10000000); fb();
        ASSERT_FALSE(fb.RawButton, 'Demarrage tenu ne simule aucun appui');
        ASSERT_EQ(fb.RawX, 5000, 'Demarrage tenu neutre');
ADVANCE_TIME(10000000); fb();
        ASSERT_FALSE(fb.RawButton, 'Demarrage tenu ne simule aucun appui');
        ASSERT_EQ(fb.RawX, 5000, 'Demarrage tenu neutre');
ADVANCE_TIME(10000000); fb();
        ASSERT_FALSE(fb.RawButton, 'Demarrage tenu ne simule aucun appui');
        ASSERT_EQ(fb.RawX, 5000, 'Demarrage tenu neutre');
ADVANCE_TIME(10000000); fb();
        ASSERT_FALSE(fb.RawButton, 'Demarrage tenu ne simule aucun appui');
        ASSERT_EQ(fb.RawX, 5000, 'Demarrage tenu neutre');
ADVANCE_TIME(10000000); fb();
        ASSERT_FALSE(fb.RawButton, 'Demarrage tenu ne simule aucun appui');
        ASSERT_EQ(fb.RawX, 5000, 'Demarrage tenu neutre');
ADVANCE_TIME(10000000); fb();
        ASSERT_FALSE(fb.RawButton, 'Demarrage tenu ne simule aucun appui');
        ASSERT_EQ(fb.RawX, 5000, 'Demarrage tenu neutre');
ADVANCE_TIME(10000000); fb();
        ASSERT_FALSE(fb.RawButton, 'Demarrage tenu ne simule aucun appui');
        ASSERT_EQ(fb.RawX, 5000, 'Demarrage tenu neutre');
ADVANCE_TIME(10000000); fb();
        ASSERT_FALSE(fb.RawButton, 'Demarrage tenu ne simule aucun appui');
        ASSERT_EQ(fb.RawX, 5000, 'Demarrage tenu neutre');
ADVANCE_TIME(10000000); fb();
        ASSERT_FALSE(fb.RawButton, 'Demarrage tenu ne simule aucun appui');
        ASSERT_EQ(fb.RawX, 5000, 'Demarrage tenu neutre');
ADVANCE_TIME(10000000); fb();
        ASSERT_FALSE(fb.RawButton, 'Demarrage tenu ne simule aucun appui');
        ASSERT_EQ(fb.RawX, 5000, 'Demarrage tenu neutre');
ADVANCE_TIME(10000000); fb();
        ASSERT_FALSE(fb.RawButton, 'Demarrage tenu ne simule aucun appui');
        ASSERT_EQ(fb.RawX, 5000, 'Demarrage tenu neutre');
ADVANCE_TIME(10000000); fb();
        ASSERT_FALSE(fb.RawButton, 'Demarrage tenu ne simule aucun appui');
        ASSERT_EQ(fb.RawX, 5000, 'Demarrage tenu neutre');
ADVANCE_TIME(10000000); fb();
        ASSERT_FALSE(fb.RawButton, 'Demarrage tenu ne simule aucun appui');
        ASSERT_EQ(fb.RawX, 5000, 'Demarrage tenu neutre');
ADVANCE_TIME(10000000); fb();
        ASSERT_FALSE(fb.RawButton, 'Demarrage tenu ne simule aucun appui');
        ASSERT_EQ(fb.RawX, 5000, 'Demarrage tenu neutre');
ADVANCE_TIME(10000000); fb();
        ASSERT_FALSE(fb.RawButton, 'Demarrage tenu ne simule aucun appui');
        ASSERT_EQ(fb.RawX, 5000, 'Demarrage tenu neutre');
ADVANCE_TIME(10000000); fb();
        ASSERT_FALSE(fb.RawButton, 'Demarrage tenu ne simule aucun appui');
        ASSERT_EQ(fb.RawX, 5000, 'Demarrage tenu neutre');
ADVANCE_TIME(10000000); fb();
        ASSERT_FALSE(fb.RawButton, 'Demarrage tenu ne simule aucun appui');
        ASSERT_EQ(fb.RawX, 5000, 'Demarrage tenu neutre');
ADVANCE_TIME(10000000); fb();
        ASSERT_FALSE(fb.RawButton, 'Demarrage tenu ne simule aucun appui');
        ASSERT_EQ(fb.RawX, 5000, 'Demarrage tenu neutre');
ADVANCE_TIME(10000000); fb();
        ASSERT_FALSE(fb.RawButton, 'Demarrage tenu ne simule aucun appui');
        ASSERT_EQ(fb.RawX, 5000, 'Demarrage tenu neutre');
ADVANCE_TIME(10000000); fb();
        ASSERT_FALSE(fb.RawButton, 'Demarrage tenu ne simule aucun appui');
        ASSERT_EQ(fb.RawX, 5000, 'Demarrage tenu neutre');
ADVANCE_TIME(10000000); fb();
        ASSERT_FALSE(fb.RawButton, 'Demarrage tenu ne simule aucun appui');
        ASSERT_EQ(fb.RawX, 5000, 'Demarrage tenu neutre');
ADVANCE_TIME(10000000); fb();
        ASSERT_FALSE(fb.RawButton, 'Demarrage tenu ne simule aucun appui');
        ASSERT_EQ(fb.RawX, 5000, 'Demarrage tenu neutre');
ADVANCE_TIME(10000000); fb();
        ASSERT_FALSE(fb.RawButton, 'Demarrage tenu ne simule aucun appui');
        ASSERT_EQ(fb.RawX, 5000, 'Demarrage tenu neutre');
ADVANCE_TIME(10000000); fb();
        ASSERT_FALSE(fb.RawButton, 'Demarrage tenu ne simule aucun appui');
        ASSERT_EQ(fb.RawX, 5000, 'Demarrage tenu neutre');
ADVANCE_TIME(10000000); fb();
        ASSERT_FALSE(fb.RawButton, 'Demarrage tenu ne simule aucun appui');
        ASSERT_EQ(fb.RawX, 5000, 'Demarrage tenu neutre');
ADVANCE_TIME(10000000); fb();
        ASSERT_FALSE(fb.RawButton, 'Demarrage tenu ne simule aucun appui');
        ASSERT_EQ(fb.RawX, 5000, 'Demarrage tenu neutre');
ADVANCE_TIME(10000000); fb();
        ASSERT_FALSE(fb.RawButton, 'Demarrage tenu ne simule aucun appui');
        ASSERT_EQ(fb.RawX, 5000, 'Demarrage tenu neutre');
ADVANCE_TIME(10000000); fb();
        ASSERT_FALSE(fb.RawButton, 'Demarrage tenu ne simule aucun appui');
        ASSERT_EQ(fb.RawX, 5000, 'Demarrage tenu neutre');
ADVANCE_TIME(10000000); fb();
        ASSERT_FALSE(fb.RawButton, 'Demarrage tenu ne simule aucun appui');
        ASSERT_EQ(fb.RawX, 5000, 'Demarrage tenu neutre');
ADVANCE_TIME(10000000); fb();
        ASSERT_FALSE(fb.RawButton, 'Demarrage tenu ne simule aucun appui');
        ASSERT_EQ(fb.RawX, 5000, 'Demarrage tenu neutre');
ADVANCE_TIME(10000000); fb();
        ASSERT_FALSE(fb.RawButton, 'Demarrage tenu ne simule aucun appui');
        ASSERT_EQ(fb.RawX, 5000, 'Demarrage tenu neutre');
ADVANCE_TIME(10000000); fb();
        ASSERT_FALSE(fb.RawButton, 'Demarrage tenu ne simule aucun appui');
        ASSERT_EQ(fb.RawX, 5000, 'Demarrage tenu neutre');
ADVANCE_TIME(10000000); fb();
        ASSERT_FALSE(fb.RawButton, 'Demarrage tenu ne simule aucun appui');
        ASSERT_EQ(fb.RawX, 5000, 'Demarrage tenu neutre');
ADVANCE_TIME(10000000); fb();
        ASSERT_FALSE(fb.RawButton, 'Demarrage tenu ne simule aucun appui');
        ASSERT_EQ(fb.RawX, 5000, 'Demarrage tenu neutre');
ADVANCE_TIME(10000000); fb();
        ASSERT_FALSE(fb.RawButton, 'Demarrage tenu ne simule aucun appui');
        ASSERT_EQ(fb.RawX, 5000, 'Demarrage tenu neutre');
ADVANCE_TIME(10000000); fb();
        ASSERT_FALSE(fb.RawButton, 'Demarrage tenu ne simule aucun appui');
        ASSERT_EQ(fb.RawX, 5000, 'Demarrage tenu neutre');
ADVANCE_TIME(10000000); fb();
        ASSERT_FALSE(fb.RawButton, 'Demarrage tenu ne simule aucun appui');
        ASSERT_EQ(fb.RawX, 5000, 'Demarrage tenu neutre');
ADVANCE_TIME(10000000); fb();
        ASSERT_FALSE(fb.RawButton, 'Demarrage tenu ne simule aucun appui');
        ASSERT_EQ(fb.RawX, 5000, 'Demarrage tenu neutre');
ADVANCE_TIME(10000000); fb();
        ASSERT_FALSE(fb.RawButton, 'Demarrage tenu ne simule aucun appui');
        ASSERT_EQ(fb.RawX, 5000, 'Demarrage tenu neutre');
ADVANCE_TIME(10000000); fb();
        ASSERT_FALSE(fb.RawButton, 'Demarrage tenu ne simule aucun appui');
        ASSERT_EQ(fb.RawX, 5000, 'Demarrage tenu neutre');
ADVANCE_TIME(10000000); fb();
        ASSERT_FALSE(fb.RawButton, 'Demarrage tenu ne simule aucun appui');
        ASSERT_EQ(fb.RawX, 5000, 'Demarrage tenu neutre');
ADVANCE_TIME(10000000); fb();
        ASSERT_FALSE(fb.RawButton, 'Demarrage tenu ne simule aucun appui');
        ASSERT_EQ(fb.RawX, 5000, 'Demarrage tenu neutre');
ADVANCE_TIME(10000000); fb();
        ASSERT_FALSE(fb.RawButton, 'Demarrage tenu ne simule aucun appui');
        ASSERT_EQ(fb.RawX, 5000, 'Demarrage tenu neutre');
ADVANCE_TIME(10000000); fb();
        ASSERT_FALSE(fb.RawButton, 'Demarrage tenu ne simule aucun appui');
        ASSERT_EQ(fb.RawX, 5000, 'Demarrage tenu neutre');
ADVANCE_TIME(10000000); fb();
        ASSERT_FALSE(fb.RawButton, 'Demarrage tenu ne simule aucun appui');
        ASSERT_EQ(fb.RawX, 5000, 'Demarrage tenu neutre');
ADVANCE_TIME(10000000); fb();
        ASSERT_FALSE(fb.RawButton, 'Demarrage tenu ne simule aucun appui');
        ASSERT_EQ(fb.RawX, 5000, 'Demarrage tenu neutre');
ADVANCE_TIME(10000000); fb();
        ASSERT_FALSE(fb.RawButton, 'Demarrage tenu ne simule aucun appui');
        ASSERT_EQ(fb.RawX, 5000, 'Demarrage tenu neutre');
ADVANCE_TIME(10000000); fb();
        ASSERT_FALSE(fb.RawButton, 'Demarrage tenu ne simule aucun appui');
        ASSERT_EQ(fb.RawX, 5000, 'Demarrage tenu neutre');
ADVANCE_TIME(10000000); fb();
        ASSERT_FALSE(fb.RawButton, 'Demarrage tenu ne simule aucun appui');
        ASSERT_EQ(fb.RawX, 5000, 'Demarrage tenu neutre');
ADVANCE_TIME(10000000); fb();
        ASSERT_FALSE(fb.RawButton, 'Demarrage tenu ne simule aucun appui');
        ASSERT_EQ(fb.RawX, 5000, 'Demarrage tenu neutre');
ADVANCE_TIME(10000000); fb();
        ASSERT_FALSE(fb.RawButton, 'Demarrage tenu ne simule aucun appui');
        ASSERT_EQ(fb.RawX, 5000, 'Demarrage tenu neutre');
ADVANCE_TIME(10000000); fb();
        ASSERT_FALSE(fb.RawButton, 'Demarrage tenu ne simule aucun appui');
        ASSERT_EQ(fb.RawX, 5000, 'Demarrage tenu neutre');
ADVANCE_TIME(10000000); fb();
        ASSERT_FALSE(fb.RawButton, 'Demarrage tenu ne simule aucun appui');
        ASSERT_EQ(fb.RawX, 5000, 'Demarrage tenu neutre');
ADVANCE_TIME(10000000); fb();
        ASSERT_FALSE(fb.RawButton, 'Demarrage tenu ne simule aucun appui');
        ASSERT_EQ(fb.RawX, 5000, 'Demarrage tenu neutre');
ADVANCE_TIME(10000000); fb();
        ASSERT_FALSE(fb.RawButton, 'Demarrage tenu ne simule aucun appui');
        ASSERT_EQ(fb.RawX, 5000, 'Demarrage tenu neutre');
ADVANCE_TIME(10000000); fb();
        ASSERT_FALSE(fb.RawButton, 'Demarrage tenu ne simule aucun appui');
        ASSERT_EQ(fb.RawX, 5000, 'Demarrage tenu neutre');
ADVANCE_TIME(10000000); fb();
        ASSERT_FALSE(fb.RawButton, 'Demarrage tenu ne simule aucun appui');
        ASSERT_EQ(fb.RawX, 5000, 'Demarrage tenu neutre');
ADVANCE_TIME(10000000); fb();
        ASSERT_FALSE(fb.RawButton, 'Demarrage tenu ne simule aucun appui');
        ASSERT_EQ(fb.RawX, 5000, 'Demarrage tenu neutre');
ADVANCE_TIME(10000000); fb();
        ASSERT_FALSE(fb.RawButton, 'Demarrage tenu ne simule aucun appui');
        ASSERT_EQ(fb.RawX, 5000, 'Demarrage tenu neutre');
ADVANCE_TIME(10000000); fb();
        ASSERT_FALSE(fb.RawButton, 'Demarrage tenu ne simule aucun appui');
        ASSERT_EQ(fb.RawX, 5000, 'Demarrage tenu neutre');
ADVANCE_TIME(10000000); fb();
        ASSERT_FALSE(fb.RawButton, 'Demarrage tenu ne simule aucun appui');
        ASSERT_EQ(fb.RawX, 5000, 'Demarrage tenu neutre');
    fb.BtnRight_Fwd_MAINT := FALSE; fb();
    fb.BtnRight_Fwd_MAINT := TRUE; fb();
    ASSERT_TRUE(fb.RawButton, 'Nouvel appui accepte');
    fb.Enable := FALSE; fb(); fb.Enable := TRUE;
    ADVANCE_TIME(10000000); fb();
        ASSERT_FALSE(fb.RawButton, 'Pas de reprise OFF ON tenu');
ADVANCE_TIME(10000000); fb();
        ASSERT_FALSE(fb.RawButton, 'Pas de reprise OFF ON tenu');
ADVANCE_TIME(10000000); fb();
        ASSERT_FALSE(fb.RawButton, 'Pas de reprise OFF ON tenu');
ADVANCE_TIME(10000000); fb();
        ASSERT_FALSE(fb.RawButton, 'Pas de reprise OFF ON tenu');
ADVANCE_TIME(10000000); fb();
        ASSERT_FALSE(fb.RawButton, 'Pas de reprise OFF ON tenu');
ADVANCE_TIME(10000000); fb();
        ASSERT_FALSE(fb.RawButton, 'Pas de reprise OFF ON tenu');
ADVANCE_TIME(10000000); fb();
        ASSERT_FALSE(fb.RawButton, 'Pas de reprise OFF ON tenu');
ADVANCE_TIME(10000000); fb();
        ASSERT_FALSE(fb.RawButton, 'Pas de reprise OFF ON tenu');
ADVANCE_TIME(10000000); fb();
        ASSERT_FALSE(fb.RawButton, 'Pas de reprise OFF ON tenu');
ADVANCE_TIME(10000000); fb();
        ASSERT_FALSE(fb.RawButton, 'Pas de reprise OFF ON tenu');
ADVANCE_TIME(10000000); fb();
        ASSERT_FALSE(fb.RawButton, 'Pas de reprise OFF ON tenu');
ADVANCE_TIME(10000000); fb();
        ASSERT_FALSE(fb.RawButton, 'Pas de reprise OFF ON tenu');
ADVANCE_TIME(10000000); fb();
        ASSERT_FALSE(fb.RawButton, 'Pas de reprise OFF ON tenu');
ADVANCE_TIME(10000000); fb();
        ASSERT_FALSE(fb.RawButton, 'Pas de reprise OFF ON tenu');
ADVANCE_TIME(10000000); fb();
        ASSERT_FALSE(fb.RawButton, 'Pas de reprise OFF ON tenu');
ADVANCE_TIME(10000000); fb();
        ASSERT_FALSE(fb.RawButton, 'Pas de reprise OFF ON tenu');
ADVANCE_TIME(10000000); fb();
        ASSERT_FALSE(fb.RawButton, 'Pas de reprise OFF ON tenu');
ADVANCE_TIME(10000000); fb();
        ASSERT_FALSE(fb.RawButton, 'Pas de reprise OFF ON tenu');
ADVANCE_TIME(10000000); fb();
        ASSERT_FALSE(fb.RawButton, 'Pas de reprise OFF ON tenu');
ADVANCE_TIME(10000000); fb();
        ASSERT_FALSE(fb.RawButton, 'Pas de reprise OFF ON tenu');
ADVANCE_TIME(10000000); fb();
        ASSERT_FALSE(fb.RawButton, 'Pas de reprise OFF ON tenu');
ADVANCE_TIME(10000000); fb();
        ASSERT_FALSE(fb.RawButton, 'Pas de reprise OFF ON tenu');
ADVANCE_TIME(10000000); fb();
        ASSERT_FALSE(fb.RawButton, 'Pas de reprise OFF ON tenu');
ADVANCE_TIME(10000000); fb();
        ASSERT_FALSE(fb.RawButton, 'Pas de reprise OFF ON tenu');
ADVANCE_TIME(10000000); fb();
        ASSERT_FALSE(fb.RawButton, 'Pas de reprise OFF ON tenu');
ADVANCE_TIME(10000000); fb();
        ASSERT_FALSE(fb.RawButton, 'Pas de reprise OFF ON tenu');
ADVANCE_TIME(10000000); fb();
        ASSERT_FALSE(fb.RawButton, 'Pas de reprise OFF ON tenu');
ADVANCE_TIME(10000000); fb();
        ASSERT_FALSE(fb.RawButton, 'Pas de reprise OFF ON tenu');
ADVANCE_TIME(10000000); fb();
        ASSERT_FALSE(fb.RawButton, 'Pas de reprise OFF ON tenu');
ADVANCE_TIME(10000000); fb();
        ASSERT_FALSE(fb.RawButton, 'Pas de reprise OFF ON tenu');
ADVANCE_TIME(10000000); fb();
        ASSERT_FALSE(fb.RawButton, 'Pas de reprise OFF ON tenu');
ADVANCE_TIME(10000000); fb();
        ASSERT_FALSE(fb.RawButton, 'Pas de reprise OFF ON tenu');
ADVANCE_TIME(10000000); fb();
        ASSERT_FALSE(fb.RawButton, 'Pas de reprise OFF ON tenu');
ADVANCE_TIME(10000000); fb();
        ASSERT_FALSE(fb.RawButton, 'Pas de reprise OFF ON tenu');
ADVANCE_TIME(10000000); fb();
        ASSERT_FALSE(fb.RawButton, 'Pas de reprise OFF ON tenu');
ADVANCE_TIME(10000000); fb();
        ASSERT_FALSE(fb.RawButton, 'Pas de reprise OFF ON tenu');
ADVANCE_TIME(10000000); fb();
        ASSERT_FALSE(fb.RawButton, 'Pas de reprise OFF ON tenu');
ADVANCE_TIME(10000000); fb();
        ASSERT_FALSE(fb.RawButton, 'Pas de reprise OFF ON tenu');
ADVANCE_TIME(10000000); fb();
        ASSERT_FALSE(fb.RawButton, 'Pas de reprise OFF ON tenu');
ADVANCE_TIME(10000000); fb();
        ASSERT_FALSE(fb.RawButton, 'Pas de reprise OFF ON tenu');
ADVANCE_TIME(10000000); fb();
        ASSERT_FALSE(fb.RawButton, 'Pas de reprise OFF ON tenu');
ADVANCE_TIME(10000000); fb();
        ASSERT_FALSE(fb.RawButton, 'Pas de reprise OFF ON tenu');
ADVANCE_TIME(10000000); fb();
        ASSERT_FALSE(fb.RawButton, 'Pas de reprise OFF ON tenu');
ADVANCE_TIME(10000000); fb();
        ASSERT_FALSE(fb.RawButton, 'Pas de reprise OFF ON tenu');
ADVANCE_TIME(10000000); fb();
        ASSERT_FALSE(fb.RawButton, 'Pas de reprise OFF ON tenu');
ADVANCE_TIME(10000000); fb();
        ASSERT_FALSE(fb.RawButton, 'Pas de reprise OFF ON tenu');
ADVANCE_TIME(10000000); fb();
        ASSERT_FALSE(fb.RawButton, 'Pas de reprise OFF ON tenu');
ADVANCE_TIME(10000000); fb();
        ASSERT_FALSE(fb.RawButton, 'Pas de reprise OFF ON tenu');
ADVANCE_TIME(10000000); fb();
        ASSERT_FALSE(fb.RawButton, 'Pas de reprise OFF ON tenu');
ADVANCE_TIME(10000000); fb();
        ASSERT_FALSE(fb.RawButton, 'Pas de reprise OFF ON tenu');
ADVANCE_TIME(10000000); fb();
        ASSERT_FALSE(fb.RawButton, 'Pas de reprise OFF ON tenu');
ADVANCE_TIME(10000000); fb();
        ASSERT_FALSE(fb.RawButton, 'Pas de reprise OFF ON tenu');
ADVANCE_TIME(10000000); fb();
        ASSERT_FALSE(fb.RawButton, 'Pas de reprise OFF ON tenu');
ADVANCE_TIME(10000000); fb();
        ASSERT_FALSE(fb.RawButton, 'Pas de reprise OFF ON tenu');
ADVANCE_TIME(10000000); fb();
        ASSERT_FALSE(fb.RawButton, 'Pas de reprise OFF ON tenu');
ADVANCE_TIME(10000000); fb();
        ASSERT_FALSE(fb.RawButton, 'Pas de reprise OFF ON tenu');
ADVANCE_TIME(10000000); fb();
        ASSERT_FALSE(fb.RawButton, 'Pas de reprise OFF ON tenu');
ADVANCE_TIME(10000000); fb();
        ASSERT_FALSE(fb.RawButton, 'Pas de reprise OFF ON tenu');
ADVANCE_TIME(10000000); fb();
        ASSERT_FALSE(fb.RawButton, 'Pas de reprise OFF ON tenu');
ADVANCE_TIME(10000000); fb();
        ASSERT_FALSE(fb.RawButton, 'Pas de reprise OFF ON tenu');
ADVANCE_TIME(10000000); fb();
        ASSERT_FALSE(fb.RawButton, 'Pas de reprise OFF ON tenu');
ADVANCE_TIME(10000000); fb();
        ASSERT_FALSE(fb.RawButton, 'Pas de reprise OFF ON tenu');
ADVANCE_TIME(10000000); fb();
        ASSERT_FALSE(fb.RawButton, 'Pas de reprise OFF ON tenu');
ADVANCE_TIME(10000000); fb();
        ASSERT_FALSE(fb.RawButton, 'Pas de reprise OFF ON tenu');
ADVANCE_TIME(10000000); fb();
        ASSERT_FALSE(fb.RawButton, 'Pas de reprise OFF ON tenu');
ADVANCE_TIME(10000000); fb();
        ASSERT_FALSE(fb.RawButton, 'Pas de reprise OFF ON tenu');
ADVANCE_TIME(10000000); fb();
        ASSERT_FALSE(fb.RawButton, 'Pas de reprise OFF ON tenu');
ADVANCE_TIME(10000000); fb();
        ASSERT_FALSE(fb.RawButton, 'Pas de reprise OFF ON tenu');
ADVANCE_TIME(10000000); fb();
        ASSERT_FALSE(fb.RawButton, 'Pas de reprise OFF ON tenu');
ADVANCE_TIME(10000000); fb();
        ASSERT_FALSE(fb.RawButton, 'Pas de reprise OFF ON tenu');
END_TEST

TEST 'TC-T418-003 Annulation avant fin maintien et conflit pendant armement'
VAR
    fb : FB_Sim_Joystick;
    i : INT;
END_VAR
    fb.Enable := TRUE; fb(); fb.BtnRight_Fwd_MAINT := TRUE; fb();
    ADVANCE_TIME(10000000); fb();
ADVANCE_TIME(10000000); fb();
ADVANCE_TIME(10000000); fb();
ADVANCE_TIME(10000000); fb();
ADVANCE_TIME(10000000); fb();
ADVANCE_TIME(10000000); fb();
ADVANCE_TIME(10000000); fb();
ADVANCE_TIME(10000000); fb();
ADVANCE_TIME(10000000); fb();
ADVANCE_TIME(10000000); fb();
ADVANCE_TIME(10000000); fb();
ADVANCE_TIME(10000000); fb();
ADVANCE_TIME(10000000); fb();
ADVANCE_TIME(10000000); fb();
ADVANCE_TIME(10000000); fb();
ADVANCE_TIME(10000000); fb();
ADVANCE_TIME(10000000); fb();
ADVANCE_TIME(10000000); fb();
ADVANCE_TIME(10000000); fb();
    fb.BtnRight_Fwd_MAINT := FALSE;
    ADVANCE_TIME(10000000); fb();
        ASSERT_EQ(fb.RawX, 5000, 'Annulation a 190 ms sans mouvement differe');
        ASSERT_FALSE(fb.RawButton, 'Appui annule');
ADVANCE_TIME(10000000); fb();
        ASSERT_EQ(fb.RawX, 5000, 'Annulation a 190 ms sans mouvement differe');
        ASSERT_FALSE(fb.RawButton, 'Appui annule');
ADVANCE_TIME(10000000); fb();
        ASSERT_EQ(fb.RawX, 5000, 'Annulation a 190 ms sans mouvement differe');
        ASSERT_FALSE(fb.RawButton, 'Appui annule');
ADVANCE_TIME(10000000); fb();
        ASSERT_EQ(fb.RawX, 5000, 'Annulation a 190 ms sans mouvement differe');
        ASSERT_FALSE(fb.RawButton, 'Appui annule');
ADVANCE_TIME(10000000); fb();
        ASSERT_EQ(fb.RawX, 5000, 'Annulation a 190 ms sans mouvement differe');
        ASSERT_FALSE(fb.RawButton, 'Appui annule');
ADVANCE_TIME(10000000); fb();
        ASSERT_EQ(fb.RawX, 5000, 'Annulation a 190 ms sans mouvement differe');
        ASSERT_FALSE(fb.RawButton, 'Appui annule');
ADVANCE_TIME(10000000); fb();
        ASSERT_EQ(fb.RawX, 5000, 'Annulation a 190 ms sans mouvement differe');
        ASSERT_FALSE(fb.RawButton, 'Appui annule');
ADVANCE_TIME(10000000); fb();
        ASSERT_EQ(fb.RawX, 5000, 'Annulation a 190 ms sans mouvement differe');
        ASSERT_FALSE(fb.RawButton, 'Appui annule');
ADVANCE_TIME(10000000); fb();
        ASSERT_EQ(fb.RawX, 5000, 'Annulation a 190 ms sans mouvement differe');
        ASSERT_FALSE(fb.RawButton, 'Appui annule');
ADVANCE_TIME(10000000); fb();
        ASSERT_EQ(fb.RawX, 5000, 'Annulation a 190 ms sans mouvement differe');
        ASSERT_FALSE(fb.RawButton, 'Appui annule');
ADVANCE_TIME(10000000); fb();
        ASSERT_EQ(fb.RawX, 5000, 'Annulation a 190 ms sans mouvement differe');
        ASSERT_FALSE(fb.RawButton, 'Appui annule');
ADVANCE_TIME(10000000); fb();
        ASSERT_EQ(fb.RawX, 5000, 'Annulation a 190 ms sans mouvement differe');
        ASSERT_FALSE(fb.RawButton, 'Appui annule');
ADVANCE_TIME(10000000); fb();
        ASSERT_EQ(fb.RawX, 5000, 'Annulation a 190 ms sans mouvement differe');
        ASSERT_FALSE(fb.RawButton, 'Appui annule');
ADVANCE_TIME(10000000); fb();
        ASSERT_EQ(fb.RawX, 5000, 'Annulation a 190 ms sans mouvement differe');
        ASSERT_FALSE(fb.RawButton, 'Appui annule');
ADVANCE_TIME(10000000); fb();
        ASSERT_EQ(fb.RawX, 5000, 'Annulation a 190 ms sans mouvement differe');
        ASSERT_FALSE(fb.RawButton, 'Appui annule');
ADVANCE_TIME(10000000); fb();
        ASSERT_EQ(fb.RawX, 5000, 'Annulation a 190 ms sans mouvement differe');
        ASSERT_FALSE(fb.RawButton, 'Appui annule');
ADVANCE_TIME(10000000); fb();
        ASSERT_EQ(fb.RawX, 5000, 'Annulation a 190 ms sans mouvement differe');
        ASSERT_FALSE(fb.RawButton, 'Appui annule');
ADVANCE_TIME(10000000); fb();
        ASSERT_EQ(fb.RawX, 5000, 'Annulation a 190 ms sans mouvement differe');
        ASSERT_FALSE(fb.RawButton, 'Appui annule');
ADVANCE_TIME(10000000); fb();
        ASSERT_EQ(fb.RawX, 5000, 'Annulation a 190 ms sans mouvement differe');
        ASSERT_FALSE(fb.RawButton, 'Appui annule');
ADVANCE_TIME(10000000); fb();
        ASSERT_EQ(fb.RawX, 5000, 'Annulation a 190 ms sans mouvement differe');
        ASSERT_FALSE(fb.RawButton, 'Appui annule');
ADVANCE_TIME(10000000); fb();
        ASSERT_EQ(fb.RawX, 5000, 'Annulation a 190 ms sans mouvement differe');
        ASSERT_FALSE(fb.RawButton, 'Appui annule');
ADVANCE_TIME(10000000); fb();
        ASSERT_EQ(fb.RawX, 5000, 'Annulation a 190 ms sans mouvement differe');
        ASSERT_FALSE(fb.RawButton, 'Appui annule');
ADVANCE_TIME(10000000); fb();
        ASSERT_EQ(fb.RawX, 5000, 'Annulation a 190 ms sans mouvement differe');
        ASSERT_FALSE(fb.RawButton, 'Appui annule');
ADVANCE_TIME(10000000); fb();
        ASSERT_EQ(fb.RawX, 5000, 'Annulation a 190 ms sans mouvement differe');
        ASSERT_FALSE(fb.RawButton, 'Appui annule');
ADVANCE_TIME(10000000); fb();
        ASSERT_EQ(fb.RawX, 5000, 'Annulation a 190 ms sans mouvement differe');
        ASSERT_FALSE(fb.RawButton, 'Appui annule');
ADVANCE_TIME(10000000); fb();
        ASSERT_EQ(fb.RawX, 5000, 'Annulation a 190 ms sans mouvement differe');
        ASSERT_FALSE(fb.RawButton, 'Appui annule');
ADVANCE_TIME(10000000); fb();
        ASSERT_EQ(fb.RawX, 5000, 'Annulation a 190 ms sans mouvement differe');
        ASSERT_FALSE(fb.RawButton, 'Appui annule');
ADVANCE_TIME(10000000); fb();
        ASSERT_EQ(fb.RawX, 5000, 'Annulation a 190 ms sans mouvement differe');
        ASSERT_FALSE(fb.RawButton, 'Appui annule');
ADVANCE_TIME(10000000); fb();
        ASSERT_EQ(fb.RawX, 5000, 'Annulation a 190 ms sans mouvement differe');
        ASSERT_FALSE(fb.RawButton, 'Appui annule');
ADVANCE_TIME(10000000); fb();
        ASSERT_EQ(fb.RawX, 5000, 'Annulation a 190 ms sans mouvement differe');
        ASSERT_FALSE(fb.RawButton, 'Appui annule');
ADVANCE_TIME(10000000); fb();
        ASSERT_EQ(fb.RawX, 5000, 'Annulation a 190 ms sans mouvement differe');
        ASSERT_FALSE(fb.RawButton, 'Appui annule');
ADVANCE_TIME(10000000); fb();
        ASSERT_EQ(fb.RawX, 5000, 'Annulation a 190 ms sans mouvement differe');
        ASSERT_FALSE(fb.RawButton, 'Appui annule');
ADVANCE_TIME(10000000); fb();
        ASSERT_EQ(fb.RawX, 5000, 'Annulation a 190 ms sans mouvement differe');
        ASSERT_FALSE(fb.RawButton, 'Appui annule');
ADVANCE_TIME(10000000); fb();
        ASSERT_EQ(fb.RawX, 5000, 'Annulation a 190 ms sans mouvement differe');
        ASSERT_FALSE(fb.RawButton, 'Appui annule');
ADVANCE_TIME(10000000); fb();
        ASSERT_EQ(fb.RawX, 5000, 'Annulation a 190 ms sans mouvement differe');
        ASSERT_FALSE(fb.RawButton, 'Appui annule');
ADVANCE_TIME(10000000); fb();
        ASSERT_EQ(fb.RawX, 5000, 'Annulation a 190 ms sans mouvement differe');
        ASSERT_FALSE(fb.RawButton, 'Appui annule');
ADVANCE_TIME(10000000); fb();
        ASSERT_EQ(fb.RawX, 5000, 'Annulation a 190 ms sans mouvement differe');
        ASSERT_FALSE(fb.RawButton, 'Appui annule');
ADVANCE_TIME(10000000); fb();
        ASSERT_EQ(fb.RawX, 5000, 'Annulation a 190 ms sans mouvement differe');
        ASSERT_FALSE(fb.RawButton, 'Appui annule');
ADVANCE_TIME(10000000); fb();
        ASSERT_EQ(fb.RawX, 5000, 'Annulation a 190 ms sans mouvement differe');
        ASSERT_FALSE(fb.RawButton, 'Appui annule');
ADVANCE_TIME(10000000); fb();
        ASSERT_EQ(fb.RawX, 5000, 'Annulation a 190 ms sans mouvement differe');
        ASSERT_FALSE(fb.RawButton, 'Appui annule');
ADVANCE_TIME(10000000); fb();
        ASSERT_EQ(fb.RawX, 5000, 'Annulation a 190 ms sans mouvement differe');
        ASSERT_FALSE(fb.RawButton, 'Appui annule');
ADVANCE_TIME(10000000); fb();
        ASSERT_EQ(fb.RawX, 5000, 'Annulation a 190 ms sans mouvement differe');
        ASSERT_FALSE(fb.RawButton, 'Appui annule');
ADVANCE_TIME(10000000); fb();
        ASSERT_EQ(fb.RawX, 5000, 'Annulation a 190 ms sans mouvement differe');
        ASSERT_FALSE(fb.RawButton, 'Appui annule');
ADVANCE_TIME(10000000); fb();
        ASSERT_EQ(fb.RawX, 5000, 'Annulation a 190 ms sans mouvement differe');
        ASSERT_FALSE(fb.RawButton, 'Appui annule');
ADVANCE_TIME(10000000); fb();
        ASSERT_EQ(fb.RawX, 5000, 'Annulation a 190 ms sans mouvement differe');
        ASSERT_FALSE(fb.RawButton, 'Appui annule');
ADVANCE_TIME(10000000); fb();
        ASSERT_EQ(fb.RawX, 5000, 'Annulation a 190 ms sans mouvement differe');
        ASSERT_FALSE(fb.RawButton, 'Appui annule');
ADVANCE_TIME(10000000); fb();
        ASSERT_EQ(fb.RawX, 5000, 'Annulation a 190 ms sans mouvement differe');
        ASSERT_FALSE(fb.RawButton, 'Appui annule');
ADVANCE_TIME(10000000); fb();
        ASSERT_EQ(fb.RawX, 5000, 'Annulation a 190 ms sans mouvement differe');
        ASSERT_FALSE(fb.RawButton, 'Appui annule');
ADVANCE_TIME(10000000); fb();
        ASSERT_EQ(fb.RawX, 5000, 'Annulation a 190 ms sans mouvement differe');
        ASSERT_FALSE(fb.RawButton, 'Appui annule');
ADVANCE_TIME(10000000); fb();
        ASSERT_EQ(fb.RawX, 5000, 'Annulation a 190 ms sans mouvement differe');
        ASSERT_FALSE(fb.RawButton, 'Appui annule');
    fb.BtnRight_Fwd_MAINT := TRUE; fb();
    fb.BtnLeft_Rev_TREMIE := TRUE; fb();
    ASSERT_FALSE(fb.RawButton, 'Conflit annule armement');
    fb.BtnLeft_Rev_TREMIE := FALSE;
    ADVANCE_TIME(10000000); fb();
        ASSERT_FALSE(fb.RawButton, 'Retirer un seul bouton ne rearme pas');
        ASSERT_EQ(fb.RawX, 5000, 'Reste neutre');
ADVANCE_TIME(10000000); fb();
        ASSERT_FALSE(fb.RawButton, 'Retirer un seul bouton ne rearme pas');
        ASSERT_EQ(fb.RawX, 5000, 'Reste neutre');
ADVANCE_TIME(10000000); fb();
        ASSERT_FALSE(fb.RawButton, 'Retirer un seul bouton ne rearme pas');
        ASSERT_EQ(fb.RawX, 5000, 'Reste neutre');
ADVANCE_TIME(10000000); fb();
        ASSERT_FALSE(fb.RawButton, 'Retirer un seul bouton ne rearme pas');
        ASSERT_EQ(fb.RawX, 5000, 'Reste neutre');
ADVANCE_TIME(10000000); fb();
        ASSERT_FALSE(fb.RawButton, 'Retirer un seul bouton ne rearme pas');
        ASSERT_EQ(fb.RawX, 5000, 'Reste neutre');
ADVANCE_TIME(10000000); fb();
        ASSERT_FALSE(fb.RawButton, 'Retirer un seul bouton ne rearme pas');
        ASSERT_EQ(fb.RawX, 5000, 'Reste neutre');
ADVANCE_TIME(10000000); fb();
        ASSERT_FALSE(fb.RawButton, 'Retirer un seul bouton ne rearme pas');
        ASSERT_EQ(fb.RawX, 5000, 'Reste neutre');
ADVANCE_TIME(10000000); fb();
        ASSERT_FALSE(fb.RawButton, 'Retirer un seul bouton ne rearme pas');
        ASSERT_EQ(fb.RawX, 5000, 'Reste neutre');
ADVANCE_TIME(10000000); fb();
        ASSERT_FALSE(fb.RawButton, 'Retirer un seul bouton ne rearme pas');
        ASSERT_EQ(fb.RawX, 5000, 'Reste neutre');
ADVANCE_TIME(10000000); fb();
        ASSERT_FALSE(fb.RawButton, 'Retirer un seul bouton ne rearme pas');
        ASSERT_EQ(fb.RawX, 5000, 'Reste neutre');
ADVANCE_TIME(10000000); fb();
        ASSERT_FALSE(fb.RawButton, 'Retirer un seul bouton ne rearme pas');
        ASSERT_EQ(fb.RawX, 5000, 'Reste neutre');
ADVANCE_TIME(10000000); fb();
        ASSERT_FALSE(fb.RawButton, 'Retirer un seul bouton ne rearme pas');
        ASSERT_EQ(fb.RawX, 5000, 'Reste neutre');
ADVANCE_TIME(10000000); fb();
        ASSERT_FALSE(fb.RawButton, 'Retirer un seul bouton ne rearme pas');
        ASSERT_EQ(fb.RawX, 5000, 'Reste neutre');
ADVANCE_TIME(10000000); fb();
        ASSERT_FALSE(fb.RawButton, 'Retirer un seul bouton ne rearme pas');
        ASSERT_EQ(fb.RawX, 5000, 'Reste neutre');
ADVANCE_TIME(10000000); fb();
        ASSERT_FALSE(fb.RawButton, 'Retirer un seul bouton ne rearme pas');
        ASSERT_EQ(fb.RawX, 5000, 'Reste neutre');
ADVANCE_TIME(10000000); fb();
        ASSERT_FALSE(fb.RawButton, 'Retirer un seul bouton ne rearme pas');
        ASSERT_EQ(fb.RawX, 5000, 'Reste neutre');
ADVANCE_TIME(10000000); fb();
        ASSERT_FALSE(fb.RawButton, 'Retirer un seul bouton ne rearme pas');
        ASSERT_EQ(fb.RawX, 5000, 'Reste neutre');
ADVANCE_TIME(10000000); fb();
        ASSERT_FALSE(fb.RawButton, 'Retirer un seul bouton ne rearme pas');
        ASSERT_EQ(fb.RawX, 5000, 'Reste neutre');
ADVANCE_TIME(10000000); fb();
        ASSERT_FALSE(fb.RawButton, 'Retirer un seul bouton ne rearme pas');
        ASSERT_EQ(fb.RawX, 5000, 'Reste neutre');
ADVANCE_TIME(10000000); fb();
        ASSERT_FALSE(fb.RawButton, 'Retirer un seul bouton ne rearme pas');
        ASSERT_EQ(fb.RawX, 5000, 'Reste neutre');
ADVANCE_TIME(10000000); fb();
        ASSERT_FALSE(fb.RawButton, 'Retirer un seul bouton ne rearme pas');
        ASSERT_EQ(fb.RawX, 5000, 'Reste neutre');
ADVANCE_TIME(10000000); fb();
        ASSERT_FALSE(fb.RawButton, 'Retirer un seul bouton ne rearme pas');
        ASSERT_EQ(fb.RawX, 5000, 'Reste neutre');
ADVANCE_TIME(10000000); fb();
        ASSERT_FALSE(fb.RawButton, 'Retirer un seul bouton ne rearme pas');
        ASSERT_EQ(fb.RawX, 5000, 'Reste neutre');
ADVANCE_TIME(10000000); fb();
        ASSERT_FALSE(fb.RawButton, 'Retirer un seul bouton ne rearme pas');
        ASSERT_EQ(fb.RawX, 5000, 'Reste neutre');
ADVANCE_TIME(10000000); fb();
        ASSERT_FALSE(fb.RawButton, 'Retirer un seul bouton ne rearme pas');
        ASSERT_EQ(fb.RawX, 5000, 'Reste neutre');
ADVANCE_TIME(10000000); fb();
        ASSERT_FALSE(fb.RawButton, 'Retirer un seul bouton ne rearme pas');
        ASSERT_EQ(fb.RawX, 5000, 'Reste neutre');
ADVANCE_TIME(10000000); fb();
        ASSERT_FALSE(fb.RawButton, 'Retirer un seul bouton ne rearme pas');
        ASSERT_EQ(fb.RawX, 5000, 'Reste neutre');
ADVANCE_TIME(10000000); fb();
        ASSERT_FALSE(fb.RawButton, 'Retirer un seul bouton ne rearme pas');
        ASSERT_EQ(fb.RawX, 5000, 'Reste neutre');
ADVANCE_TIME(10000000); fb();
        ASSERT_FALSE(fb.RawButton, 'Retirer un seul bouton ne rearme pas');
        ASSERT_EQ(fb.RawX, 5000, 'Reste neutre');
ADVANCE_TIME(10000000); fb();
        ASSERT_FALSE(fb.RawButton, 'Retirer un seul bouton ne rearme pas');
        ASSERT_EQ(fb.RawX, 5000, 'Reste neutre');
ADVANCE_TIME(10000000); fb();
        ASSERT_FALSE(fb.RawButton, 'Retirer un seul bouton ne rearme pas');
        ASSERT_EQ(fb.RawX, 5000, 'Reste neutre');
ADVANCE_TIME(10000000); fb();
        ASSERT_FALSE(fb.RawButton, 'Retirer un seul bouton ne rearme pas');
        ASSERT_EQ(fb.RawX, 5000, 'Reste neutre');
ADVANCE_TIME(10000000); fb();
        ASSERT_FALSE(fb.RawButton, 'Retirer un seul bouton ne rearme pas');
        ASSERT_EQ(fb.RawX, 5000, 'Reste neutre');
ADVANCE_TIME(10000000); fb();
        ASSERT_FALSE(fb.RawButton, 'Retirer un seul bouton ne rearme pas');
        ASSERT_EQ(fb.RawX, 5000, 'Reste neutre');
ADVANCE_TIME(10000000); fb();
        ASSERT_FALSE(fb.RawButton, 'Retirer un seul bouton ne rearme pas');
        ASSERT_EQ(fb.RawX, 5000, 'Reste neutre');
ADVANCE_TIME(10000000); fb();
        ASSERT_FALSE(fb.RawButton, 'Retirer un seul bouton ne rearme pas');
        ASSERT_EQ(fb.RawX, 5000, 'Reste neutre');
ADVANCE_TIME(10000000); fb();
        ASSERT_FALSE(fb.RawButton, 'Retirer un seul bouton ne rearme pas');
        ASSERT_EQ(fb.RawX, 5000, 'Reste neutre');
ADVANCE_TIME(10000000); fb();
        ASSERT_FALSE(fb.RawButton, 'Retirer un seul bouton ne rearme pas');
        ASSERT_EQ(fb.RawX, 5000, 'Reste neutre');
ADVANCE_TIME(10000000); fb();
        ASSERT_FALSE(fb.RawButton, 'Retirer un seul bouton ne rearme pas');
        ASSERT_EQ(fb.RawX, 5000, 'Reste neutre');
ADVANCE_TIME(10000000); fb();
        ASSERT_FALSE(fb.RawButton, 'Retirer un seul bouton ne rearme pas');
        ASSERT_EQ(fb.RawX, 5000, 'Reste neutre');
ADVANCE_TIME(10000000); fb();
        ASSERT_FALSE(fb.RawButton, 'Retirer un seul bouton ne rearme pas');
        ASSERT_EQ(fb.RawX, 5000, 'Reste neutre');
ADVANCE_TIME(10000000); fb();
        ASSERT_FALSE(fb.RawButton, 'Retirer un seul bouton ne rearme pas');
        ASSERT_EQ(fb.RawX, 5000, 'Reste neutre');
ADVANCE_TIME(10000000); fb();
        ASSERT_FALSE(fb.RawButton, 'Retirer un seul bouton ne rearme pas');
        ASSERT_EQ(fb.RawX, 5000, 'Reste neutre');
ADVANCE_TIME(10000000); fb();
        ASSERT_FALSE(fb.RawButton, 'Retirer un seul bouton ne rearme pas');
        ASSERT_EQ(fb.RawX, 5000, 'Reste neutre');
ADVANCE_TIME(10000000); fb();
        ASSERT_FALSE(fb.RawButton, 'Retirer un seul bouton ne rearme pas');
        ASSERT_EQ(fb.RawX, 5000, 'Reste neutre');
ADVANCE_TIME(10000000); fb();
        ASSERT_FALSE(fb.RawButton, 'Retirer un seul bouton ne rearme pas');
        ASSERT_EQ(fb.RawX, 5000, 'Reste neutre');
ADVANCE_TIME(10000000); fb();
        ASSERT_FALSE(fb.RawButton, 'Retirer un seul bouton ne rearme pas');
        ASSERT_EQ(fb.RawX, 5000, 'Reste neutre');
ADVANCE_TIME(10000000); fb();
        ASSERT_FALSE(fb.RawButton, 'Retirer un seul bouton ne rearme pas');
        ASSERT_EQ(fb.RawX, 5000, 'Reste neutre');
ADVANCE_TIME(10000000); fb();
        ASSERT_FALSE(fb.RawButton, 'Retirer un seul bouton ne rearme pas');
        ASSERT_EQ(fb.RawX, 5000, 'Reste neutre');
ADVANCE_TIME(10000000); fb();
        ASSERT_FALSE(fb.RawButton, 'Retirer un seul bouton ne rearme pas');
        ASSERT_EQ(fb.RawX, 5000, 'Reste neutre');
ADVANCE_TIME(10000000); fb();
        ASSERT_FALSE(fb.RawButton, 'Retirer un seul bouton ne rearme pas');
        ASSERT_EQ(fb.RawX, 5000, 'Reste neutre');
ADVANCE_TIME(10000000); fb();
        ASSERT_FALSE(fb.RawButton, 'Retirer un seul bouton ne rearme pas');
        ASSERT_EQ(fb.RawX, 5000, 'Reste neutre');
ADVANCE_TIME(10000000); fb();
        ASSERT_FALSE(fb.RawButton, 'Retirer un seul bouton ne rearme pas');
        ASSERT_EQ(fb.RawX, 5000, 'Reste neutre');
ADVANCE_TIME(10000000); fb();
        ASSERT_FALSE(fb.RawButton, 'Retirer un seul bouton ne rearme pas');
        ASSERT_EQ(fb.RawX, 5000, 'Reste neutre');
ADVANCE_TIME(10000000); fb();
        ASSERT_FALSE(fb.RawButton, 'Retirer un seul bouton ne rearme pas');
        ASSERT_EQ(fb.RawX, 5000, 'Reste neutre');
ADVANCE_TIME(10000000); fb();
        ASSERT_FALSE(fb.RawButton, 'Retirer un seul bouton ne rearme pas');
        ASSERT_EQ(fb.RawX, 5000, 'Reste neutre');
ADVANCE_TIME(10000000); fb();
        ASSERT_FALSE(fb.RawButton, 'Retirer un seul bouton ne rearme pas');
        ASSERT_EQ(fb.RawX, 5000, 'Reste neutre');
ADVANCE_TIME(10000000); fb();
        ASSERT_FALSE(fb.RawButton, 'Retirer un seul bouton ne rearme pas');
        ASSERT_EQ(fb.RawX, 5000, 'Reste neutre');
ADVANCE_TIME(10000000); fb();
        ASSERT_FALSE(fb.RawButton, 'Retirer un seul bouton ne rearme pas');
        ASSERT_EQ(fb.RawX, 5000, 'Reste neutre');
ADVANCE_TIME(10000000); fb();
        ASSERT_FALSE(fb.RawButton, 'Retirer un seul bouton ne rearme pas');
        ASSERT_EQ(fb.RawX, 5000, 'Reste neutre');
ADVANCE_TIME(10000000); fb();
        ASSERT_FALSE(fb.RawButton, 'Retirer un seul bouton ne rearme pas');
        ASSERT_EQ(fb.RawX, 5000, 'Reste neutre');
ADVANCE_TIME(10000000); fb();
        ASSERT_FALSE(fb.RawButton, 'Retirer un seul bouton ne rearme pas');
        ASSERT_EQ(fb.RawX, 5000, 'Reste neutre');
ADVANCE_TIME(10000000); fb();
        ASSERT_FALSE(fb.RawButton, 'Retirer un seul bouton ne rearme pas');
        ASSERT_EQ(fb.RawX, 5000, 'Reste neutre');
ADVANCE_TIME(10000000); fb();
        ASSERT_FALSE(fb.RawButton, 'Retirer un seul bouton ne rearme pas');
        ASSERT_EQ(fb.RawX, 5000, 'Reste neutre');
ADVANCE_TIME(10000000); fb();
        ASSERT_FALSE(fb.RawButton, 'Retirer un seul bouton ne rearme pas');
        ASSERT_EQ(fb.RawX, 5000, 'Reste neutre');
ADVANCE_TIME(10000000); fb();
        ASSERT_FALSE(fb.RawButton, 'Retirer un seul bouton ne rearme pas');
        ASSERT_EQ(fb.RawX, 5000, 'Reste neutre');
ADVANCE_TIME(10000000); fb();
        ASSERT_FALSE(fb.RawButton, 'Retirer un seul bouton ne rearme pas');
        ASSERT_EQ(fb.RawX, 5000, 'Reste neutre');
ADVANCE_TIME(10000000); fb();
        ASSERT_FALSE(fb.RawButton, 'Retirer un seul bouton ne rearme pas');
        ASSERT_EQ(fb.RawX, 5000, 'Reste neutre');
ADVANCE_TIME(10000000); fb();
        ASSERT_FALSE(fb.RawButton, 'Retirer un seul bouton ne rearme pas');
        ASSERT_EQ(fb.RawX, 5000, 'Reste neutre');
ADVANCE_TIME(10000000); fb();
        ASSERT_FALSE(fb.RawButton, 'Retirer un seul bouton ne rearme pas');
        ASSERT_EQ(fb.RawX, 5000, 'Reste neutre');
END_TEST

TEST 'TC-T418-004 Inversion et nouvel appui pendant retour refuses'
VAR
    fb : FB_Sim_Joystick;
    i : INT;
END_VAR
    fb.Enable := TRUE; fb(); fb.BtnRight_Fwd_MAINT := TRUE;
    ADVANCE_TIME(10000000); fb();
ADVANCE_TIME(10000000); fb();
ADVANCE_TIME(10000000); fb();
ADVANCE_TIME(10000000); fb();
ADVANCE_TIME(10000000); fb();
ADVANCE_TIME(10000000); fb();
ADVANCE_TIME(10000000); fb();
ADVANCE_TIME(10000000); fb();
ADVANCE_TIME(10000000); fb();
ADVANCE_TIME(10000000); fb();
ADVANCE_TIME(10000000); fb();
ADVANCE_TIME(10000000); fb();
ADVANCE_TIME(10000000); fb();
ADVANCE_TIME(10000000); fb();
ADVANCE_TIME(10000000); fb();
ADVANCE_TIME(10000000); fb();
ADVANCE_TIME(10000000); fb();
ADVANCE_TIME(10000000); fb();
ADVANCE_TIME(10000000); fb();
ADVANCE_TIME(10000000); fb();
ADVANCE_TIME(10000000); fb();
ADVANCE_TIME(10000000); fb();
ADVANCE_TIME(10000000); fb();
ADVANCE_TIME(10000000); fb();
ADVANCE_TIME(10000000); fb();
ADVANCE_TIME(10000000); fb();
ADVANCE_TIME(10000000); fb();
ADVANCE_TIME(10000000); fb();
ADVANCE_TIME(10000000); fb();
ADVANCE_TIME(10000000); fb();
ADVANCE_TIME(10000000); fb();
ADVANCE_TIME(10000000); fb();
ADVANCE_TIME(10000000); fb();
ADVANCE_TIME(10000000); fb();
ADVANCE_TIME(10000000); fb();
ADVANCE_TIME(10000000); fb();
ADVANCE_TIME(10000000); fb();
ADVANCE_TIME(10000000); fb();
ADVANCE_TIME(10000000); fb();
ADVANCE_TIME(10000000); fb();
ADVANCE_TIME(10000000); fb();
ADVANCE_TIME(10000000); fb();
ADVANCE_TIME(10000000); fb();
ADVANCE_TIME(10000000); fb();
ADVANCE_TIME(10000000); fb();
ADVANCE_TIME(10000000); fb();
ADVANCE_TIME(10000000); fb();
ADVANCE_TIME(10000000); fb();
ADVANCE_TIME(10000000); fb();
ADVANCE_TIME(10000000); fb();
ADVANCE_TIME(10000000); fb();
ADVANCE_TIME(10000000); fb();
ADVANCE_TIME(10000000); fb();
ADVANCE_TIME(10000000); fb();
ADVANCE_TIME(10000000); fb();
ADVANCE_TIME(10000000); fb();
ADVANCE_TIME(10000000); fb();
ADVANCE_TIME(10000000); fb();
ADVANCE_TIME(10000000); fb();
ADVANCE_TIME(10000000); fb();
ADVANCE_TIME(10000000); fb();
ADVANCE_TIME(10000000); fb();
ADVANCE_TIME(10000000); fb();
ADVANCE_TIME(10000000); fb();
ADVANCE_TIME(10000000); fb();
ADVANCE_TIME(10000000); fb();
ADVANCE_TIME(10000000); fb();
ADVANCE_TIME(10000000); fb();
ADVANCE_TIME(10000000); fb();
ADVANCE_TIME(10000000); fb();
ADVANCE_TIME(10000000); fb();
ADVANCE_TIME(10000000); fb();
ADVANCE_TIME(10000000); fb();
ADVANCE_TIME(10000000); fb();
ADVANCE_TIME(10000000); fb();
ADVANCE_TIME(10000000); fb();
ADVANCE_TIME(10000000); fb();
ADVANCE_TIME(10000000); fb();
ADVANCE_TIME(10000000); fb();
ADVANCE_TIME(10000000); fb();
ADVANCE_TIME(10000000); fb();
ADVANCE_TIME(10000000); fb();
ADVANCE_TIME(10000000); fb();
ADVANCE_TIME(10000000); fb();
ADVANCE_TIME(10000000); fb();
ADVANCE_TIME(10000000); fb();
ADVANCE_TIME(10000000); fb();
ADVANCE_TIME(10000000); fb();
ADVANCE_TIME(10000000); fb();
ADVANCE_TIME(10000000); fb();
ADVANCE_TIME(10000000); fb();
ADVANCE_TIME(10000000); fb();
ADVANCE_TIME(10000000); fb();
ADVANCE_TIME(10000000); fb();
ADVANCE_TIME(10000000); fb();
ADVANCE_TIME(10000000); fb();
ADVANCE_TIME(10000000); fb();
ADVANCE_TIME(10000000); fb();
ADVANCE_TIME(10000000); fb();
ADVANCE_TIME(10000000); fb();
ADVANCE_TIME(10000000); fb();
ADVANCE_TIME(10000000); fb();
ADVANCE_TIME(10000000); fb();
ADVANCE_TIME(10000000); fb();
ADVANCE_TIME(10000000); fb();
ADVANCE_TIME(10000000); fb();
ADVANCE_TIME(10000000); fb();
ADVANCE_TIME(10000000); fb();
ADVANCE_TIME(10000000); fb();
ADVANCE_TIME(10000000); fb();
ADVANCE_TIME(10000000); fb();
ADVANCE_TIME(10000000); fb();
ADVANCE_TIME(10000000); fb();
ADVANCE_TIME(10000000); fb();
ADVANCE_TIME(10000000); fb();
ADVANCE_TIME(10000000); fb();
ADVANCE_TIME(10000000); fb();
ADVANCE_TIME(10000000); fb();
ADVANCE_TIME(10000000); fb();
ADVANCE_TIME(10000000); fb();
ADVANCE_TIME(10000000); fb();
ADVANCE_TIME(10000000); fb();
ADVANCE_TIME(10000000); fb();
ADVANCE_TIME(10000000); fb();
ADVANCE_TIME(10000000); fb();
ADVANCE_TIME(10000000); fb();
ADVANCE_TIME(10000000); fb();
ADVANCE_TIME(10000000); fb();
ADVANCE_TIME(10000000); fb();
ADVANCE_TIME(10000000); fb();
ADVANCE_TIME(10000000); fb();
ADVANCE_TIME(10000000); fb();
ADVANCE_TIME(10000000); fb();
ADVANCE_TIME(10000000); fb();
ADVANCE_TIME(10000000); fb();
ADVANCE_TIME(10000000); fb();
ADVANCE_TIME(10000000); fb();
ADVANCE_TIME(10000000); fb();
ADVANCE_TIME(10000000); fb();
ADVANCE_TIME(10000000); fb();
ADVANCE_TIME(10000000); fb();
ADVANCE_TIME(10000000); fb();
ADVANCE_TIME(10000000); fb();
ADVANCE_TIME(10000000); fb();
ADVANCE_TIME(10000000); fb();
ADVANCE_TIME(10000000); fb();
ADVANCE_TIME(10000000); fb();
ADVANCE_TIME(10000000); fb();
ADVANCE_TIME(10000000); fb();
ADVANCE_TIME(10000000); fb();
ADVANCE_TIME(10000000); fb();
ADVANCE_TIME(10000000); fb();
ADVANCE_TIME(10000000); fb();
ADVANCE_TIME(10000000); fb();
ADVANCE_TIME(10000000); fb();
ADVANCE_TIME(10000000); fb();
ADVANCE_TIME(10000000); fb();
ADVANCE_TIME(10000000); fb();
ADVANCE_TIME(10000000); fb();
ADVANCE_TIME(10000000); fb();
ADVANCE_TIME(10000000); fb();
ADVANCE_TIME(10000000); fb();
ADVANCE_TIME(10000000); fb();
ADVANCE_TIME(10000000); fb();
ADVANCE_TIME(10000000); fb();
ADVANCE_TIME(10000000); fb();
ADVANCE_TIME(10000000); fb();
ADVANCE_TIME(10000000); fb();
ADVANCE_TIME(10000000); fb();
ADVANCE_TIME(10000000); fb();
ADVANCE_TIME(10000000); fb();
ADVANCE_TIME(10000000); fb();
ADVANCE_TIME(10000000); fb();
ADVANCE_TIME(10000000); fb();
ADVANCE_TIME(10000000); fb();
ADVANCE_TIME(10000000); fb();
ADVANCE_TIME(10000000); fb();
ADVANCE_TIME(10000000); fb();
ADVANCE_TIME(10000000); fb();
ADVANCE_TIME(10000000); fb();
    ASSERT_TRUE(fb.RawX > 9000, 'Geste initial effectif');
    fb.BtnRight_Fwd_MAINT := FALSE; fb.BtnLeft_Rev_TREMIE := TRUE;
    ADVANCE_TIME(10000000); fb();
        ASSERT_TRUE(fb.RawX >= 5000, 'Inversion directe ne franchit pas le neutre');
        ASSERT_FALSE(fb.RawButton, 'Inversion ne rearme pas');
ADVANCE_TIME(10000000); fb();
        ASSERT_TRUE(fb.RawX >= 5000, 'Inversion directe ne franchit pas le neutre');
        ASSERT_FALSE(fb.RawButton, 'Inversion ne rearme pas');
ADVANCE_TIME(10000000); fb();
        ASSERT_TRUE(fb.RawX >= 5000, 'Inversion directe ne franchit pas le neutre');
        ASSERT_FALSE(fb.RawButton, 'Inversion ne rearme pas');
ADVANCE_TIME(10000000); fb();
        ASSERT_TRUE(fb.RawX >= 5000, 'Inversion directe ne franchit pas le neutre');
        ASSERT_FALSE(fb.RawButton, 'Inversion ne rearme pas');
ADVANCE_TIME(10000000); fb();
        ASSERT_TRUE(fb.RawX >= 5000, 'Inversion directe ne franchit pas le neutre');
        ASSERT_FALSE(fb.RawButton, 'Inversion ne rearme pas');
ADVANCE_TIME(10000000); fb();
        ASSERT_TRUE(fb.RawX >= 5000, 'Inversion directe ne franchit pas le neutre');
        ASSERT_FALSE(fb.RawButton, 'Inversion ne rearme pas');
ADVANCE_TIME(10000000); fb();
        ASSERT_TRUE(fb.RawX >= 5000, 'Inversion directe ne franchit pas le neutre');
        ASSERT_FALSE(fb.RawButton, 'Inversion ne rearme pas');
ADVANCE_TIME(10000000); fb();
        ASSERT_TRUE(fb.RawX >= 5000, 'Inversion directe ne franchit pas le neutre');
        ASSERT_FALSE(fb.RawButton, 'Inversion ne rearme pas');
ADVANCE_TIME(10000000); fb();
        ASSERT_TRUE(fb.RawX >= 5000, 'Inversion directe ne franchit pas le neutre');
        ASSERT_FALSE(fb.RawButton, 'Inversion ne rearme pas');
ADVANCE_TIME(10000000); fb();
        ASSERT_TRUE(fb.RawX >= 5000, 'Inversion directe ne franchit pas le neutre');
        ASSERT_FALSE(fb.RawButton, 'Inversion ne rearme pas');
ADVANCE_TIME(10000000); fb();
        ASSERT_TRUE(fb.RawX >= 5000, 'Inversion directe ne franchit pas le neutre');
        ASSERT_FALSE(fb.RawButton, 'Inversion ne rearme pas');
ADVANCE_TIME(10000000); fb();
        ASSERT_TRUE(fb.RawX >= 5000, 'Inversion directe ne franchit pas le neutre');
        ASSERT_FALSE(fb.RawButton, 'Inversion ne rearme pas');
ADVANCE_TIME(10000000); fb();
        ASSERT_TRUE(fb.RawX >= 5000, 'Inversion directe ne franchit pas le neutre');
        ASSERT_FALSE(fb.RawButton, 'Inversion ne rearme pas');
ADVANCE_TIME(10000000); fb();
        ASSERT_TRUE(fb.RawX >= 5000, 'Inversion directe ne franchit pas le neutre');
        ASSERT_FALSE(fb.RawButton, 'Inversion ne rearme pas');
ADVANCE_TIME(10000000); fb();
        ASSERT_TRUE(fb.RawX >= 5000, 'Inversion directe ne franchit pas le neutre');
        ASSERT_FALSE(fb.RawButton, 'Inversion ne rearme pas');
ADVANCE_TIME(10000000); fb();
        ASSERT_TRUE(fb.RawX >= 5000, 'Inversion directe ne franchit pas le neutre');
        ASSERT_FALSE(fb.RawButton, 'Inversion ne rearme pas');
ADVANCE_TIME(10000000); fb();
        ASSERT_TRUE(fb.RawX >= 5000, 'Inversion directe ne franchit pas le neutre');
        ASSERT_FALSE(fb.RawButton, 'Inversion ne rearme pas');
ADVANCE_TIME(10000000); fb();
        ASSERT_TRUE(fb.RawX >= 5000, 'Inversion directe ne franchit pas le neutre');
        ASSERT_FALSE(fb.RawButton, 'Inversion ne rearme pas');
ADVANCE_TIME(10000000); fb();
        ASSERT_TRUE(fb.RawX >= 5000, 'Inversion directe ne franchit pas le neutre');
        ASSERT_FALSE(fb.RawButton, 'Inversion ne rearme pas');
ADVANCE_TIME(10000000); fb();
        ASSERT_TRUE(fb.RawX >= 5000, 'Inversion directe ne franchit pas le neutre');
        ASSERT_FALSE(fb.RawButton, 'Inversion ne rearme pas');
ADVANCE_TIME(10000000); fb();
        ASSERT_TRUE(fb.RawX >= 5000, 'Inversion directe ne franchit pas le neutre');
        ASSERT_FALSE(fb.RawButton, 'Inversion ne rearme pas');
ADVANCE_TIME(10000000); fb();
        ASSERT_TRUE(fb.RawX >= 5000, 'Inversion directe ne franchit pas le neutre');
        ASSERT_FALSE(fb.RawButton, 'Inversion ne rearme pas');
ADVANCE_TIME(10000000); fb();
        ASSERT_TRUE(fb.RawX >= 5000, 'Inversion directe ne franchit pas le neutre');
        ASSERT_FALSE(fb.RawButton, 'Inversion ne rearme pas');
ADVANCE_TIME(10000000); fb();
        ASSERT_TRUE(fb.RawX >= 5000, 'Inversion directe ne franchit pas le neutre');
        ASSERT_FALSE(fb.RawButton, 'Inversion ne rearme pas');
ADVANCE_TIME(10000000); fb();
        ASSERT_TRUE(fb.RawX >= 5000, 'Inversion directe ne franchit pas le neutre');
        ASSERT_FALSE(fb.RawButton, 'Inversion ne rearme pas');
ADVANCE_TIME(10000000); fb();
        ASSERT_TRUE(fb.RawX >= 5000, 'Inversion directe ne franchit pas le neutre');
        ASSERT_FALSE(fb.RawButton, 'Inversion ne rearme pas');
ADVANCE_TIME(10000000); fb();
        ASSERT_TRUE(fb.RawX >= 5000, 'Inversion directe ne franchit pas le neutre');
        ASSERT_FALSE(fb.RawButton, 'Inversion ne rearme pas');
ADVANCE_TIME(10000000); fb();
        ASSERT_TRUE(fb.RawX >= 5000, 'Inversion directe ne franchit pas le neutre');
        ASSERT_FALSE(fb.RawButton, 'Inversion ne rearme pas');
ADVANCE_TIME(10000000); fb();
        ASSERT_TRUE(fb.RawX >= 5000, 'Inversion directe ne franchit pas le neutre');
        ASSERT_FALSE(fb.RawButton, 'Inversion ne rearme pas');
ADVANCE_TIME(10000000); fb();
        ASSERT_TRUE(fb.RawX >= 5000, 'Inversion directe ne franchit pas le neutre');
        ASSERT_FALSE(fb.RawButton, 'Inversion ne rearme pas');
ADVANCE_TIME(10000000); fb();
        ASSERT_TRUE(fb.RawX >= 5000, 'Inversion directe ne franchit pas le neutre');
        ASSERT_FALSE(fb.RawButton, 'Inversion ne rearme pas');
ADVANCE_TIME(10000000); fb();
        ASSERT_TRUE(fb.RawX >= 5000, 'Inversion directe ne franchit pas le neutre');
        ASSERT_FALSE(fb.RawButton, 'Inversion ne rearme pas');
ADVANCE_TIME(10000000); fb();
        ASSERT_TRUE(fb.RawX >= 5000, 'Inversion directe ne franchit pas le neutre');
        ASSERT_FALSE(fb.RawButton, 'Inversion ne rearme pas');
ADVANCE_TIME(10000000); fb();
        ASSERT_TRUE(fb.RawX >= 5000, 'Inversion directe ne franchit pas le neutre');
        ASSERT_FALSE(fb.RawButton, 'Inversion ne rearme pas');
ADVANCE_TIME(10000000); fb();
        ASSERT_TRUE(fb.RawX >= 5000, 'Inversion directe ne franchit pas le neutre');
        ASSERT_FALSE(fb.RawButton, 'Inversion ne rearme pas');
ADVANCE_TIME(10000000); fb();
        ASSERT_TRUE(fb.RawX >= 5000, 'Inversion directe ne franchit pas le neutre');
        ASSERT_FALSE(fb.RawButton, 'Inversion ne rearme pas');
ADVANCE_TIME(10000000); fb();
        ASSERT_TRUE(fb.RawX >= 5000, 'Inversion directe ne franchit pas le neutre');
        ASSERT_FALSE(fb.RawButton, 'Inversion ne rearme pas');
ADVANCE_TIME(10000000); fb();
        ASSERT_TRUE(fb.RawX >= 5000, 'Inversion directe ne franchit pas le neutre');
        ASSERT_FALSE(fb.RawButton, 'Inversion ne rearme pas');
ADVANCE_TIME(10000000); fb();
        ASSERT_TRUE(fb.RawX >= 5000, 'Inversion directe ne franchit pas le neutre');
        ASSERT_FALSE(fb.RawButton, 'Inversion ne rearme pas');
ADVANCE_TIME(10000000); fb();
        ASSERT_TRUE(fb.RawX >= 5000, 'Inversion directe ne franchit pas le neutre');
        ASSERT_FALSE(fb.RawButton, 'Inversion ne rearme pas');
ADVANCE_TIME(10000000); fb();
        ASSERT_TRUE(fb.RawX >= 5000, 'Inversion directe ne franchit pas le neutre');
        ASSERT_FALSE(fb.RawButton, 'Inversion ne rearme pas');
ADVANCE_TIME(10000000); fb();
        ASSERT_TRUE(fb.RawX >= 5000, 'Inversion directe ne franchit pas le neutre');
        ASSERT_FALSE(fb.RawButton, 'Inversion ne rearme pas');
ADVANCE_TIME(10000000); fb();
        ASSERT_TRUE(fb.RawX >= 5000, 'Inversion directe ne franchit pas le neutre');
        ASSERT_FALSE(fb.RawButton, 'Inversion ne rearme pas');
ADVANCE_TIME(10000000); fb();
        ASSERT_TRUE(fb.RawX >= 5000, 'Inversion directe ne franchit pas le neutre');
        ASSERT_FALSE(fb.RawButton, 'Inversion ne rearme pas');
ADVANCE_TIME(10000000); fb();
        ASSERT_TRUE(fb.RawX >= 5000, 'Inversion directe ne franchit pas le neutre');
        ASSERT_FALSE(fb.RawButton, 'Inversion ne rearme pas');
ADVANCE_TIME(10000000); fb();
        ASSERT_TRUE(fb.RawX >= 5000, 'Inversion directe ne franchit pas le neutre');
        ASSERT_FALSE(fb.RawButton, 'Inversion ne rearme pas');
ADVANCE_TIME(10000000); fb();
        ASSERT_TRUE(fb.RawX >= 5000, 'Inversion directe ne franchit pas le neutre');
        ASSERT_FALSE(fb.RawButton, 'Inversion ne rearme pas');
ADVANCE_TIME(10000000); fb();
        ASSERT_TRUE(fb.RawX >= 5000, 'Inversion directe ne franchit pas le neutre');
        ASSERT_FALSE(fb.RawButton, 'Inversion ne rearme pas');
ADVANCE_TIME(10000000); fb();
        ASSERT_TRUE(fb.RawX >= 5000, 'Inversion directe ne franchit pas le neutre');
        ASSERT_FALSE(fb.RawButton, 'Inversion ne rearme pas');
ADVANCE_TIME(10000000); fb();
        ASSERT_TRUE(fb.RawX >= 5000, 'Inversion directe ne franchit pas le neutre');
        ASSERT_FALSE(fb.RawButton, 'Inversion ne rearme pas');
ADVANCE_TIME(10000000); fb();
        ASSERT_TRUE(fb.RawX >= 5000, 'Inversion directe ne franchit pas le neutre');
        ASSERT_FALSE(fb.RawButton, 'Inversion ne rearme pas');
ADVANCE_TIME(10000000); fb();
        ASSERT_TRUE(fb.RawX >= 5000, 'Inversion directe ne franchit pas le neutre');
        ASSERT_FALSE(fb.RawButton, 'Inversion ne rearme pas');
ADVANCE_TIME(10000000); fb();
        ASSERT_TRUE(fb.RawX >= 5000, 'Inversion directe ne franchit pas le neutre');
        ASSERT_FALSE(fb.RawButton, 'Inversion ne rearme pas');
ADVANCE_TIME(10000000); fb();
        ASSERT_TRUE(fb.RawX >= 5000, 'Inversion directe ne franchit pas le neutre');
        ASSERT_FALSE(fb.RawButton, 'Inversion ne rearme pas');
ADVANCE_TIME(10000000); fb();
        ASSERT_TRUE(fb.RawX >= 5000, 'Inversion directe ne franchit pas le neutre');
        ASSERT_FALSE(fb.RawButton, 'Inversion ne rearme pas');
ADVANCE_TIME(10000000); fb();
        ASSERT_TRUE(fb.RawX >= 5000, 'Inversion directe ne franchit pas le neutre');
        ASSERT_FALSE(fb.RawButton, 'Inversion ne rearme pas');
ADVANCE_TIME(10000000); fb();
        ASSERT_TRUE(fb.RawX >= 5000, 'Inversion directe ne franchit pas le neutre');
        ASSERT_FALSE(fb.RawButton, 'Inversion ne rearme pas');
ADVANCE_TIME(10000000); fb();
        ASSERT_TRUE(fb.RawX >= 5000, 'Inversion directe ne franchit pas le neutre');
        ASSERT_FALSE(fb.RawButton, 'Inversion ne rearme pas');
ADVANCE_TIME(10000000); fb();
        ASSERT_TRUE(fb.RawX >= 5000, 'Inversion directe ne franchit pas le neutre');
        ASSERT_FALSE(fb.RawButton, 'Inversion ne rearme pas');
ADVANCE_TIME(10000000); fb();
        ASSERT_TRUE(fb.RawX >= 5000, 'Inversion directe ne franchit pas le neutre');
        ASSERT_FALSE(fb.RawButton, 'Inversion ne rearme pas');
    fb.BtnLeft_Rev_TREMIE := FALSE; fb();
    fb.BtnRight_Fwd_MAINT := TRUE;
    ADVANCE_TIME(10000000); fb();
ADVANCE_TIME(10000000); fb();
ADVANCE_TIME(10000000); fb();
ADVANCE_TIME(10000000); fb();
ADVANCE_TIME(10000000); fb();
ADVANCE_TIME(10000000); fb();
ADVANCE_TIME(10000000); fb();
ADVANCE_TIME(10000000); fb();
ADVANCE_TIME(10000000); fb();
ADVANCE_TIME(10000000); fb();
ADVANCE_TIME(10000000); fb();
ADVANCE_TIME(10000000); fb();
ADVANCE_TIME(10000000); fb();
ADVANCE_TIME(10000000); fb();
ADVANCE_TIME(10000000); fb();
ADVANCE_TIME(10000000); fb();
ADVANCE_TIME(10000000); fb();
ADVANCE_TIME(10000000); fb();
ADVANCE_TIME(10000000); fb();
ADVANCE_TIME(10000000); fb();
ADVANCE_TIME(10000000); fb();
ADVANCE_TIME(10000000); fb();
ADVANCE_TIME(10000000); fb();
ADVANCE_TIME(10000000); fb();
ADVANCE_TIME(10000000); fb();
ADVANCE_TIME(10000000); fb();
ADVANCE_TIME(10000000); fb();
ADVANCE_TIME(10000000); fb();
ADVANCE_TIME(10000000); fb();
ADVANCE_TIME(10000000); fb();
ADVANCE_TIME(10000000); fb();
ADVANCE_TIME(10000000); fb();
ADVANCE_TIME(10000000); fb();
ADVANCE_TIME(10000000); fb();
ADVANCE_TIME(10000000); fb();
ADVANCE_TIME(10000000); fb();
ADVANCE_TIME(10000000); fb();
ADVANCE_TIME(10000000); fb();
ADVANCE_TIME(10000000); fb();
ADVANCE_TIME(10000000); fb();
ADVANCE_TIME(10000000); fb();
ADVANCE_TIME(10000000); fb();
ADVANCE_TIME(10000000); fb();
ADVANCE_TIME(10000000); fb();
ADVANCE_TIME(10000000); fb();
ADVANCE_TIME(10000000); fb();
ADVANCE_TIME(10000000); fb();
ADVANCE_TIME(10000000); fb();
ADVANCE_TIME(10000000); fb();
ADVANCE_TIME(10000000); fb();
ADVANCE_TIME(10000000); fb();
ADVANCE_TIME(10000000); fb();
ADVANCE_TIME(10000000); fb();
ADVANCE_TIME(10000000); fb();
ADVANCE_TIME(10000000); fb();
ADVANCE_TIME(10000000); fb();
ADVANCE_TIME(10000000); fb();
ADVANCE_TIME(10000000); fb();
ADVANCE_TIME(10000000); fb();
ADVANCE_TIME(10000000); fb();
ADVANCE_TIME(10000000); fb();
ADVANCE_TIME(10000000); fb();
ADVANCE_TIME(10000000); fb();
ADVANCE_TIME(10000000); fb();
ADVANCE_TIME(10000000); fb();
ADVANCE_TIME(10000000); fb();
ADVANCE_TIME(10000000); fb();
ADVANCE_TIME(10000000); fb();
ADVANCE_TIME(10000000); fb();
ADVANCE_TIME(10000000); fb();
ADVANCE_TIME(10000000); fb();
ADVANCE_TIME(10000000); fb();
ADVANCE_TIME(10000000); fb();
ADVANCE_TIME(10000000); fb();
ADVANCE_TIME(10000000); fb();
ADVANCE_TIME(10000000); fb();
ADVANCE_TIME(10000000); fb();
ADVANCE_TIME(10000000); fb();
ADVANCE_TIME(10000000); fb();
ADVANCE_TIME(10000000); fb();
ADVANCE_TIME(10000000); fb();
ADVANCE_TIME(10000000); fb();
ADVANCE_TIME(10000000); fb();
ADVANCE_TIME(10000000); fb();
ADVANCE_TIME(10000000); fb();
ADVANCE_TIME(10000000); fb();
ADVANCE_TIME(10000000); fb();
ADVANCE_TIME(10000000); fb();
ADVANCE_TIME(10000000); fb();
ADVANCE_TIME(10000000); fb();
ADVANCE_TIME(10000000); fb();
ADVANCE_TIME(10000000); fb();
ADVANCE_TIME(10000000); fb();
ADVANCE_TIME(10000000); fb();
ADVANCE_TIME(10000000); fb();
ADVANCE_TIME(10000000); fb();
ADVANCE_TIME(10000000); fb();
ADVANCE_TIME(10000000); fb();
ADVANCE_TIME(10000000); fb();
ADVANCE_TIME(10000000); fb();
    fb.BtnRight_Fwd_MAINT := FALSE; fb();
    fb.BtnLeft_Rev_TREMIE := TRUE;
    ADVANCE_TIME(10000000); fb();
        ASSERT_FALSE(fb.RawButton, 'Appui pendant retour non mis en attente');
        ASSERT_TRUE(fb.RawX >= 5000, 'Pas de depart inverse differe');
ADVANCE_TIME(10000000); fb();
        ASSERT_FALSE(fb.RawButton, 'Appui pendant retour non mis en attente');
        ASSERT_TRUE(fb.RawX >= 5000, 'Pas de depart inverse differe');
ADVANCE_TIME(10000000); fb();
        ASSERT_FALSE(fb.RawButton, 'Appui pendant retour non mis en attente');
        ASSERT_TRUE(fb.RawX >= 5000, 'Pas de depart inverse differe');
ADVANCE_TIME(10000000); fb();
        ASSERT_FALSE(fb.RawButton, 'Appui pendant retour non mis en attente');
        ASSERT_TRUE(fb.RawX >= 5000, 'Pas de depart inverse differe');
ADVANCE_TIME(10000000); fb();
        ASSERT_FALSE(fb.RawButton, 'Appui pendant retour non mis en attente');
        ASSERT_TRUE(fb.RawX >= 5000, 'Pas de depart inverse differe');
ADVANCE_TIME(10000000); fb();
        ASSERT_FALSE(fb.RawButton, 'Appui pendant retour non mis en attente');
        ASSERT_TRUE(fb.RawX >= 5000, 'Pas de depart inverse differe');
ADVANCE_TIME(10000000); fb();
        ASSERT_FALSE(fb.RawButton, 'Appui pendant retour non mis en attente');
        ASSERT_TRUE(fb.RawX >= 5000, 'Pas de depart inverse differe');
ADVANCE_TIME(10000000); fb();
        ASSERT_FALSE(fb.RawButton, 'Appui pendant retour non mis en attente');
        ASSERT_TRUE(fb.RawX >= 5000, 'Pas de depart inverse differe');
ADVANCE_TIME(10000000); fb();
        ASSERT_FALSE(fb.RawButton, 'Appui pendant retour non mis en attente');
        ASSERT_TRUE(fb.RawX >= 5000, 'Pas de depart inverse differe');
ADVANCE_TIME(10000000); fb();
        ASSERT_FALSE(fb.RawButton, 'Appui pendant retour non mis en attente');
        ASSERT_TRUE(fb.RawX >= 5000, 'Pas de depart inverse differe');
ADVANCE_TIME(10000000); fb();
        ASSERT_FALSE(fb.RawButton, 'Appui pendant retour non mis en attente');
        ASSERT_TRUE(fb.RawX >= 5000, 'Pas de depart inverse differe');
ADVANCE_TIME(10000000); fb();
        ASSERT_FALSE(fb.RawButton, 'Appui pendant retour non mis en attente');
        ASSERT_TRUE(fb.RawX >= 5000, 'Pas de depart inverse differe');
ADVANCE_TIME(10000000); fb();
        ASSERT_FALSE(fb.RawButton, 'Appui pendant retour non mis en attente');
        ASSERT_TRUE(fb.RawX >= 5000, 'Pas de depart inverse differe');
ADVANCE_TIME(10000000); fb();
        ASSERT_FALSE(fb.RawButton, 'Appui pendant retour non mis en attente');
        ASSERT_TRUE(fb.RawX >= 5000, 'Pas de depart inverse differe');
ADVANCE_TIME(10000000); fb();
        ASSERT_FALSE(fb.RawButton, 'Appui pendant retour non mis en attente');
        ASSERT_TRUE(fb.RawX >= 5000, 'Pas de depart inverse differe');
ADVANCE_TIME(10000000); fb();
        ASSERT_FALSE(fb.RawButton, 'Appui pendant retour non mis en attente');
        ASSERT_TRUE(fb.RawX >= 5000, 'Pas de depart inverse differe');
ADVANCE_TIME(10000000); fb();
        ASSERT_FALSE(fb.RawButton, 'Appui pendant retour non mis en attente');
        ASSERT_TRUE(fb.RawX >= 5000, 'Pas de depart inverse differe');
ADVANCE_TIME(10000000); fb();
        ASSERT_FALSE(fb.RawButton, 'Appui pendant retour non mis en attente');
        ASSERT_TRUE(fb.RawX >= 5000, 'Pas de depart inverse differe');
ADVANCE_TIME(10000000); fb();
        ASSERT_FALSE(fb.RawButton, 'Appui pendant retour non mis en attente');
        ASSERT_TRUE(fb.RawX >= 5000, 'Pas de depart inverse differe');
ADVANCE_TIME(10000000); fb();
        ASSERT_FALSE(fb.RawButton, 'Appui pendant retour non mis en attente');
        ASSERT_TRUE(fb.RawX >= 5000, 'Pas de depart inverse differe');
ADVANCE_TIME(10000000); fb();
        ASSERT_FALSE(fb.RawButton, 'Appui pendant retour non mis en attente');
        ASSERT_TRUE(fb.RawX >= 5000, 'Pas de depart inverse differe');
ADVANCE_TIME(10000000); fb();
        ASSERT_FALSE(fb.RawButton, 'Appui pendant retour non mis en attente');
        ASSERT_TRUE(fb.RawX >= 5000, 'Pas de depart inverse differe');
ADVANCE_TIME(10000000); fb();
        ASSERT_FALSE(fb.RawButton, 'Appui pendant retour non mis en attente');
        ASSERT_TRUE(fb.RawX >= 5000, 'Pas de depart inverse differe');
ADVANCE_TIME(10000000); fb();
        ASSERT_FALSE(fb.RawButton, 'Appui pendant retour non mis en attente');
        ASSERT_TRUE(fb.RawX >= 5000, 'Pas de depart inverse differe');
ADVANCE_TIME(10000000); fb();
        ASSERT_FALSE(fb.RawButton, 'Appui pendant retour non mis en attente');
        ASSERT_TRUE(fb.RawX >= 5000, 'Pas de depart inverse differe');
ADVANCE_TIME(10000000); fb();
        ASSERT_FALSE(fb.RawButton, 'Appui pendant retour non mis en attente');
        ASSERT_TRUE(fb.RawX >= 5000, 'Pas de depart inverse differe');
ADVANCE_TIME(10000000); fb();
        ASSERT_FALSE(fb.RawButton, 'Appui pendant retour non mis en attente');
        ASSERT_TRUE(fb.RawX >= 5000, 'Pas de depart inverse differe');
ADVANCE_TIME(10000000); fb();
        ASSERT_FALSE(fb.RawButton, 'Appui pendant retour non mis en attente');
        ASSERT_TRUE(fb.RawX >= 5000, 'Pas de depart inverse differe');
ADVANCE_TIME(10000000); fb();
        ASSERT_FALSE(fb.RawButton, 'Appui pendant retour non mis en attente');
        ASSERT_TRUE(fb.RawX >= 5000, 'Pas de depart inverse differe');
ADVANCE_TIME(10000000); fb();
        ASSERT_FALSE(fb.RawButton, 'Appui pendant retour non mis en attente');
        ASSERT_TRUE(fb.RawX >= 5000, 'Pas de depart inverse differe');
ADVANCE_TIME(10000000); fb();
        ASSERT_FALSE(fb.RawButton, 'Appui pendant retour non mis en attente');
        ASSERT_TRUE(fb.RawX >= 5000, 'Pas de depart inverse differe');
ADVANCE_TIME(10000000); fb();
        ASSERT_FALSE(fb.RawButton, 'Appui pendant retour non mis en attente');
        ASSERT_TRUE(fb.RawX >= 5000, 'Pas de depart inverse differe');
ADVANCE_TIME(10000000); fb();
        ASSERT_FALSE(fb.RawButton, 'Appui pendant retour non mis en attente');
        ASSERT_TRUE(fb.RawX >= 5000, 'Pas de depart inverse differe');
ADVANCE_TIME(10000000); fb();
        ASSERT_FALSE(fb.RawButton, 'Appui pendant retour non mis en attente');
        ASSERT_TRUE(fb.RawX >= 5000, 'Pas de depart inverse differe');
ADVANCE_TIME(10000000); fb();
        ASSERT_FALSE(fb.RawButton, 'Appui pendant retour non mis en attente');
        ASSERT_TRUE(fb.RawX >= 5000, 'Pas de depart inverse differe');
ADVANCE_TIME(10000000); fb();
        ASSERT_FALSE(fb.RawButton, 'Appui pendant retour non mis en attente');
        ASSERT_TRUE(fb.RawX >= 5000, 'Pas de depart inverse differe');
ADVANCE_TIME(10000000); fb();
        ASSERT_FALSE(fb.RawButton, 'Appui pendant retour non mis en attente');
        ASSERT_TRUE(fb.RawX >= 5000, 'Pas de depart inverse differe');
ADVANCE_TIME(10000000); fb();
        ASSERT_FALSE(fb.RawButton, 'Appui pendant retour non mis en attente');
        ASSERT_TRUE(fb.RawX >= 5000, 'Pas de depart inverse differe');
ADVANCE_TIME(10000000); fb();
        ASSERT_FALSE(fb.RawButton, 'Appui pendant retour non mis en attente');
        ASSERT_TRUE(fb.RawX >= 5000, 'Pas de depart inverse differe');
ADVANCE_TIME(10000000); fb();
        ASSERT_FALSE(fb.RawButton, 'Appui pendant retour non mis en attente');
        ASSERT_TRUE(fb.RawX >= 5000, 'Pas de depart inverse differe');
ADVANCE_TIME(10000000); fb();
        ASSERT_FALSE(fb.RawButton, 'Appui pendant retour non mis en attente');
        ASSERT_TRUE(fb.RawX >= 5000, 'Pas de depart inverse differe');
ADVANCE_TIME(10000000); fb();
        ASSERT_FALSE(fb.RawButton, 'Appui pendant retour non mis en attente');
        ASSERT_TRUE(fb.RawX >= 5000, 'Pas de depart inverse differe');
ADVANCE_TIME(10000000); fb();
        ASSERT_FALSE(fb.RawButton, 'Appui pendant retour non mis en attente');
        ASSERT_TRUE(fb.RawX >= 5000, 'Pas de depart inverse differe');
ADVANCE_TIME(10000000); fb();
        ASSERT_FALSE(fb.RawButton, 'Appui pendant retour non mis en attente');
        ASSERT_TRUE(fb.RawX >= 5000, 'Pas de depart inverse differe');
ADVANCE_TIME(10000000); fb();
        ASSERT_FALSE(fb.RawButton, 'Appui pendant retour non mis en attente');
        ASSERT_TRUE(fb.RawX >= 5000, 'Pas de depart inverse differe');
ADVANCE_TIME(10000000); fb();
        ASSERT_FALSE(fb.RawButton, 'Appui pendant retour non mis en attente');
        ASSERT_TRUE(fb.RawX >= 5000, 'Pas de depart inverse differe');
ADVANCE_TIME(10000000); fb();
        ASSERT_FALSE(fb.RawButton, 'Appui pendant retour non mis en attente');
        ASSERT_TRUE(fb.RawX >= 5000, 'Pas de depart inverse differe');
ADVANCE_TIME(10000000); fb();
        ASSERT_FALSE(fb.RawButton, 'Appui pendant retour non mis en attente');
        ASSERT_TRUE(fb.RawX >= 5000, 'Pas de depart inverse differe');
ADVANCE_TIME(10000000); fb();
        ASSERT_FALSE(fb.RawButton, 'Appui pendant retour non mis en attente');
        ASSERT_TRUE(fb.RawX >= 5000, 'Pas de depart inverse differe');
ADVANCE_TIME(10000000); fb();
        ASSERT_FALSE(fb.RawButton, 'Appui pendant retour non mis en attente');
        ASSERT_TRUE(fb.RawX >= 5000, 'Pas de depart inverse differe');
ADVANCE_TIME(10000000); fb();
        ASSERT_FALSE(fb.RawButton, 'Appui pendant retour non mis en attente');
        ASSERT_TRUE(fb.RawX >= 5000, 'Pas de depart inverse differe');
ADVANCE_TIME(10000000); fb();
        ASSERT_FALSE(fb.RawButton, 'Appui pendant retour non mis en attente');
        ASSERT_TRUE(fb.RawX >= 5000, 'Pas de depart inverse differe');
ADVANCE_TIME(10000000); fb();
        ASSERT_FALSE(fb.RawButton, 'Appui pendant retour non mis en attente');
        ASSERT_TRUE(fb.RawX >= 5000, 'Pas de depart inverse differe');
ADVANCE_TIME(10000000); fb();
        ASSERT_FALSE(fb.RawButton, 'Appui pendant retour non mis en attente');
        ASSERT_TRUE(fb.RawX >= 5000, 'Pas de depart inverse differe');
ADVANCE_TIME(10000000); fb();
        ASSERT_FALSE(fb.RawButton, 'Appui pendant retour non mis en attente');
        ASSERT_TRUE(fb.RawX >= 5000, 'Pas de depart inverse differe');
ADVANCE_TIME(10000000); fb();
        ASSERT_FALSE(fb.RawButton, 'Appui pendant retour non mis en attente');
        ASSERT_TRUE(fb.RawX >= 5000, 'Pas de depart inverse differe');
ADVANCE_TIME(10000000); fb();
        ASSERT_FALSE(fb.RawButton, 'Appui pendant retour non mis en attente');
        ASSERT_TRUE(fb.RawX >= 5000, 'Pas de depart inverse differe');
ADVANCE_TIME(10000000); fb();
        ASSERT_FALSE(fb.RawButton, 'Appui pendant retour non mis en attente');
        ASSERT_TRUE(fb.RawX >= 5000, 'Pas de depart inverse differe');
ADVANCE_TIME(10000000); fb();
        ASSERT_FALSE(fb.RawButton, 'Appui pendant retour non mis en attente');
        ASSERT_TRUE(fb.RawX >= 5000, 'Pas de depart inverse differe');
ADVANCE_TIME(10000000); fb();
        ASSERT_FALSE(fb.RawButton, 'Appui pendant retour non mis en attente');
        ASSERT_TRUE(fb.RawX >= 5000, 'Pas de depart inverse differe');
    fb.BtnLeft_Rev_TREMIE := FALSE; fb(); fb.BtnLeft_Rev_TREMIE := TRUE;
    ADVANCE_TIME(10000000); fb();
ADVANCE_TIME(10000000); fb();
ADVANCE_TIME(10000000); fb();
ADVANCE_TIME(10000000); fb();
ADVANCE_TIME(10000000); fb();
ADVANCE_TIME(10000000); fb();
ADVANCE_TIME(10000000); fb();
ADVANCE_TIME(10000000); fb();
ADVANCE_TIME(10000000); fb();
ADVANCE_TIME(10000000); fb();
ADVANCE_TIME(10000000); fb();
ADVANCE_TIME(10000000); fb();
ADVANCE_TIME(10000000); fb();
ADVANCE_TIME(10000000); fb();
ADVANCE_TIME(10000000); fb();
ADVANCE_TIME(10000000); fb();
ADVANCE_TIME(10000000); fb();
ADVANCE_TIME(10000000); fb();
ADVANCE_TIME(10000000); fb();
ADVANCE_TIME(10000000); fb();
ADVANCE_TIME(10000000); fb();
ADVANCE_TIME(10000000); fb();
ADVANCE_TIME(10000000); fb();
ADVANCE_TIME(10000000); fb();
ADVANCE_TIME(10000000); fb();
ADVANCE_TIME(10000000); fb();
ADVANCE_TIME(10000000); fb();
ADVANCE_TIME(10000000); fb();
ADVANCE_TIME(10000000); fb();
ADVANCE_TIME(10000000); fb();
ADVANCE_TIME(10000000); fb();
ADVANCE_TIME(10000000); fb();
ADVANCE_TIME(10000000); fb();
ADVANCE_TIME(10000000); fb();
ADVANCE_TIME(10000000); fb();
ADVANCE_TIME(10000000); fb();
ADVANCE_TIME(10000000); fb();
ADVANCE_TIME(10000000); fb();
ADVANCE_TIME(10000000); fb();
ADVANCE_TIME(10000000); fb();
ADVANCE_TIME(10000000); fb();
ADVANCE_TIME(10000000); fb();
ADVANCE_TIME(10000000); fb();
ADVANCE_TIME(10000000); fb();
ADVANCE_TIME(10000000); fb();
ADVANCE_TIME(10000000); fb();
ADVANCE_TIME(10000000); fb();
ADVANCE_TIME(10000000); fb();
ADVANCE_TIME(10000000); fb();
ADVANCE_TIME(10000000); fb();
ADVANCE_TIME(10000000); fb();
ADVANCE_TIME(10000000); fb();
ADVANCE_TIME(10000000); fb();
ADVANCE_TIME(10000000); fb();
ADVANCE_TIME(10000000); fb();
ADVANCE_TIME(10000000); fb();
ADVANCE_TIME(10000000); fb();
ADVANCE_TIME(10000000); fb();
ADVANCE_TIME(10000000); fb();
ADVANCE_TIME(10000000); fb();
ADVANCE_TIME(10000000); fb();
ADVANCE_TIME(10000000); fb();
ADVANCE_TIME(10000000); fb();
ADVANCE_TIME(10000000); fb();
ADVANCE_TIME(10000000); fb();
ADVANCE_TIME(10000000); fb();
ADVANCE_TIME(10000000); fb();
ADVANCE_TIME(10000000); fb();
ADVANCE_TIME(10000000); fb();
ADVANCE_TIME(10000000); fb();
ADVANCE_TIME(10000000); fb();
ADVANCE_TIME(10000000); fb();
ADVANCE_TIME(10000000); fb();
ADVANCE_TIME(10000000); fb();
ADVANCE_TIME(10000000); fb();
ADVANCE_TIME(10000000); fb();
ADVANCE_TIME(10000000); fb();
ADVANCE_TIME(10000000); fb();
ADVANCE_TIME(10000000); fb();
ADVANCE_TIME(10000000); fb();
    ASSERT_TRUE(fb.RawX < 5000, 'Nouvel appui apres retour accepte');
END_TEST
